(* IEC 61131-3 sources: daoli-st-library/DL_Device (part 14) *)

(* ---- FB_DL_BushingDrawStartSeq.st ---- *)
// FB_DL_BushingDrawStartSeq v1.0.0
// 开源溯源：clean-room 自研（族 DL_Device，ST 生态实测 0 命中，无外部代码引入）
(*
  功能: 拉丝启动八相顺控：IDLE→HEAT→(达标保持300s)DRIP→(检滴料)ATTACH→(丝根附着)RAMP
        →(达目标速度)STEADY→(断丝)BREAK→(重接)RAMP；RAMP 按 20 m/min² 斜坡（增量 (20/60)·fCycleS）。
        联锁：①HEAT 相温度未达 fTempTarget − 5 °C 前 xWinderEnable 必须 FALSE；
              ②BREAK 相速度降至 fSpeedTarget·0.3 并保持 60 s 等重接，超时锁存；
              ③FAULT 相 xWinderEnable = FALSE 且 fSpeedCmd = 0（安全侧），仅 xReset 解除。
  邻件: 与 FC_DL_BushingTempZoneCalc（分区温度）、FC_DL_BushingPowerBalanceCalc（功率平衡）同族，本件不调用 FC。
  码表: 9331 入参非有限｜9332 组态非法(fCycleS/fTempTarget/fSpeedTarget≤0)｜9333 相超时(1800/60/60/120/60 s)
        9334 相位落 ELSE 兜底｜9335 信息级进入稳态拉丝。故障码锁存至 xReset 上升沿。
  边界: 无方法块/无属性块/无全局变量/无物理 IO 地址；六 TON 单相独占且无条件刷新；速度单位统一 m/min。
*)
TYPE E_DL_DrawStartPhase :
(
    IDLE   := 0,        // 空闲：等启动指令 [-] / Idle, waiting start
    HEAT   := 10,       // 升温：漏板升到目标 − 5 °C 并保持 [-] / Heating bushing
    DRIP   := 20,       // 滴料：等玻璃液滴料 [-] / Waiting for drip
    ATTACH := 30,       // 附着：等丝根附着 [-] / Waiting for attachment
    RAMP   := 40,       // 升速：按 20 m/min² 升至目标 [-] / Ramping up
    STEADY := 50,       // 稳态：稳态拉丝 [-] / Steady drawing
    BREAK  := 60,       // 断丝：降速至 30% 待重接 [-] / Break, slow for re-attach
    FAULT  := 90        // 故障：锁存，仅复位沿可出 [-] / Fault latched
);
END_TYPE
FUNCTION_BLOCK FB_DL_BushingDrawStartSeq
VAR_INPUT
    xEnable         : BOOL := FALSE;    // 使能，FALSE 时冻结在 IDLE [-] / Enable gate
    xStart          : BOOL := FALSE;    // 启动指令，上升沿有效 [-] / Start rising edge
    xReset          : BOOL := FALSE;    // 复位，上升沿清故障锁存 [-] / Reset rising edge
    fBushingTemp    : REAL := 25.0;     // 漏板实测温度 [°C] / Measured bushing temperature [degC]
    fTempTarget     : REAL := 1250.0;   // 漏板目标温度 [°C]，域 > 0 / Target temperature [degC]
    xDripDetected   : BOOL := FALSE;    // 滴料检出反馈 [-] / Drip detected
    xStrandAttached : BOOL := FALSE;    // 丝根附着反馈 [-] / Strand attached
    fWinderSpeed    : REAL := 0.0;      // 卷绕实测线速 [m/min] / Measured winder speed [m/min]
    fSpeedTarget    : REAL := 900.0;    // 目标拉丝线速 [m/min]，域 > 0 / Target speed [m/min]
    xBreakDetected  : BOOL := FALSE;    // 断丝检出反馈 [-] / Break detected
    fCycleS         : REAL := 0.01;     // 任务周期 [s]，域 > 0 / Task cycle time [s]
END_VAR
VAR_OUTPUT
    ePhase        : E_DL_DrawStartPhase;    // 相位出口，段尾单点映射 [-] / Phase outlet
    xHeatEnable   : BOOL;                   // 漏板加热使能（仅 HEAT 相）[-] / Heat enable
    xWinderEnable : BOOL;                   // 卷绕使能（温度达标后）[-] / Winder enable
    fSpeedCmd     : REAL;                   // 线速指令 [m/min] / Speed command [m/min]
    xSteady       : BOOL;                   // 稳态标志（STEADY 相电平）[-] / Steady flag
    xFault        : BOOL;                   // 故障锁存标志 [-] / Fault latch flag
    uErrorId      : UDINT;                  // 事件码，0 = 无事件 / Event code
END_VAR
VAR
    tonHeat   : TON;                        // 温度达标保持窗 300 s，无条件刷新 / Temperature dwell
    tonHeatTo : TON;                        // 升温相总超时 1800 s，无条件刷新 / Heat timeout
    tonDrip   : TON;                        // 滴料相超时 60 s，无条件刷新 / Drip timeout
    tonAttach : TON;                        // 附着相超时 60 s，无条件刷新 / Attach timeout
    tonRamp   : TON;                        // 升速相超时 120 s，无条件刷新 / Ramp timeout
    tonBreak  : TON;                        // 断丝保持窗 60 s，无条件刷新 / Break hold window
    rtStart   : R_TRIG;                     // 启动沿实例，无条件刷新 / Start edge instance
    rtReset   : R_TRIG;                     // 复位沿实例，无条件刷新 / Reset edge instance
    _ePhase   : E_DL_DrawStartPhase := E_DL_DrawStartPhase.IDLE;    // 内部相位，CASE 唯一写入 / Internal phase
    _fSpeed   : REAL := 0.0;                // 速度斜坡内部量 [m/min] / Ramp speed [m/min]
    _bReady   : BOOL := FALSE;              // 温度达标判据 [-] / Temperature ready judgement
    _bFault   : BOOL := FALSE;              // 故障锁存位（锁存量，仅复位沿清）/ Latched fault bit
    _uFault   : UDINT := 16#0000;           // 故障码锁存（锁存量，仅复位沿清）/ Latched fault code
    _uInfo    : UDINT := 16#0000;           // 信息码，每拍重算 / Transient info code
END_VAR
// 段 0：定时器与沿实例无条件周期刷新（禁置于 IF/CASE 内，R7/R188）/ Unconditional refresh
rtStart(CLK := xStart);                                                     // 启动沿每拍必调 / Start edge
rtReset(CLK := xReset);                                                     // 复位沿每拍必调 / Reset edge
tonHeat(IN := (_ePhase = E_DL_DrawStartPhase.HEAT) AND (fBushingTemp >= (fTempTarget - 5.0)), PT := T#300S);
tonHeatTo(IN := (_ePhase = E_DL_DrawStartPhase.HEAT), PT := T#1800S);       // 升温总超时 / Heat timeout
tonDrip(IN := (_ePhase = E_DL_DrawStartPhase.DRIP), PT := T#60S);           // 滴料超时 / Drip timeout
tonAttach(IN := (_ePhase = E_DL_DrawStartPhase.ATTACH), PT := T#60S);       // 附着超时 / Attach timeout
tonRamp(IN := (_ePhase = E_DL_DrawStartPhase.RAMP), PT := T#120S);          // 升速超时 / Ramp timeout
tonBreak(IN := (_ePhase = E_DL_DrawStartPhase.BREAK), PT := T#60S);         // 断丝保持窗 / Break window
// 段 1：单拍量预清零（锁存量 _bFault/_uFault/_fSpeed 不入清单，R187）/ One-shot clear
_uInfo := 16#0000;                  // 信息码每拍重算 / Info code recomputed
_bReady := FALSE;                   // 温度达标判据缺省假 / Ready default false
// 段 2：非有限闸与组态域闸（归因唯一，逐因独立码，R190）/ Gate stage
IF (fBushingTemp <> fBushingTemp) OR (fTempTarget <> fTempTarget)
   OR (fWinderSpeed <> fWinderSpeed) OR (fSpeedTarget <> fSpeedTarget) OR (fCycleS <> fCycleS)
   OR (ABS(fBushingTemp) >= 3.0E38) OR (ABS(fTempTarget) >= 3.0E38)
   OR (ABS(fWinderSpeed) >= 3.0E38) OR (ABS(fSpeedTarget) >= 3.0E38) OR (ABS(fCycleS) >= 3.0E38) THEN
    _uFault := 16#0002_9331;        // 故障级：入参非有限 / Fault: non-finite input
    _bFault := TRUE;                // 置故障锁存（R45 配对）/ Set fault latch
END_IF
IF (fCycleS <= 1.0E-6) OR (fTempTarget <= 1.0E-6) OR (fSpeedTarget <= 1.0E-6) THEN
    _uFault := 16#0002_9332;        // 故障级：组态非法 / Fault: illegal configuration
    _bFault := TRUE;                // 置故障锁存（R45 配对）/ Set fault latch
END_IF
// 段 3：温度达标判据（HEAT 与 DRIP 共用，禁 EQUAL 比较）/ Temperature ready judgement
IF fBushingTemp >= (fTempTarget - 5.0) THEN
    _bReady := TRUE;                // 达目标 − 5 °C / Reached target minus margin
END_IF
// 段 4：复位沿（FAULT 唯一解除路径）/ Reset edge, only exit from fault
IF rtReset.Q THEN                   // rtReset.Q = 当拍量 / Reset edge per scan
    IF _ePhase = E_DL_DrawStartPhase.FAULT THEN
        _ePhase := E_DL_DrawStartPhase.IDLE;    // 故障相迁出回空闲 / Fault exits to idle
    END_IF
    _fSpeed := 0.0;                 // 斜坡量归零（锁存量解除）/ Ramp cleared on reset
    _bFault := FALSE;               // 清故障锁存位（仅此解除沿可清）/ Clear latched bit
    _uFault := 16#0000;             // 清故障锁存码（仅此解除沿可清）/ Clear latched code
END_IF
// 段 5：相位机（本拍合法事件优先于超时，R275）/ Phase machine
CASE _ePhase OF
E_DL_DrawStartPhase.IDLE:
    IF _bFault THEN
        _ePhase := E_DL_DrawStartPhase.FAULT;       // 聚合故障进故障相 / Enter fault
    ELSIF rtStart.Q AND xEnable THEN
        _fSpeed := 0.0;                             // 启动前进度清零 / Ramp reset on start
        _ePhase := E_DL_DrawStartPhase.HEAT;        // 进升温相 / Enter heat
    END_IF
E_DL_DrawStartPhase.HEAT:
    IF _bFault THEN
        _ePhase := E_DL_DrawStartPhase.FAULT;       // 故障优先 / Fault first
    ELSIF NOT xEnable THEN
        _ePhase := E_DL_DrawStartPhase.IDLE;        // 使能撤销回空闲 / Enable dropped
    ELSIF tonHeat.Q THEN
        _ePhase := E_DL_DrawStartPhase.DRIP;        // 达标保持 300 s：进滴料相 / Dwell done, drip
    ELSIF tonHeatTo.Q THEN
        _uFault := 16#0002_9333;                    // 故障级：升温相超时 / Heat timeout
        _bFault := TRUE;                            // 置故障锁存（R45 配对）/ Set latch
        _ePhase := E_DL_DrawStartPhase.FAULT;       // 进故障相 / Enter fault
    END_IF
E_DL_DrawStartPhase.DRIP:
    IF _bFault THEN
        _ePhase := E_DL_DrawStartPhase.FAULT;       // 故障优先 / Fault first
    ELSIF NOT xEnable THEN
        _ePhase := E_DL_DrawStartPhase.IDLE;        // 使能撤销回空闲（安全侧，R92 修）/ Enable dropped to IDLE
    ELSIF xDripDetected THEN
        _ePhase := E_DL_DrawStartPhase.ATTACH;      // 检出滴料：进附着相 / Drip seen, attach
    ELSIF tonDrip.Q THEN
        _uFault := 16#0002_9333;                    // 故障级：滴料相超时 / Drip timeout
        _bFault := TRUE;                            // 置故障锁存（R45 配对）/ Set latch
        _ePhase := E_DL_DrawStartPhase.FAULT;       // 进故障相 / Enter fault
    END_IF
E_DL_DrawStartPhase.ATTACH:
    IF _bFault THEN
        _ePhase := E_DL_DrawStartPhase.FAULT;       // 故障优先 / Fault first
    ELSIF NOT xEnable THEN
        _ePhase := E_DL_DrawStartPhase.IDLE;        // 使能撤销回空闲（安全侧，R92 修）/ Enable dropped to IDLE
    ELSIF xStrandAttached THEN
        _fSpeed := 0.0;                             // 升速前进度清零 / Reset ramp before spinning
        _ePhase := E_DL_DrawStartPhase.RAMP;        // 进升速相 / Enter ramp
    ELSIF tonAttach.Q THEN
        _uFault := 16#0002_9333;                    // 故障级：附着相超时 / Attach timeout
        _bFault := TRUE;                            // 置故障锁存（R45 配对）/ Set latch
        _ePhase := E_DL_DrawStartPhase.FAULT;       // 进故障相 / Enter fault
    END_IF
E_DL_DrawStartPhase.RAMP:
    IF _bFault THEN
        _ePhase := E_DL_DrawStartPhase.FAULT;       // 故障优先 / Fault first
    ELSIF NOT xEnable THEN
        _ePhase := E_DL_DrawStartPhase.IDLE;        // 使能撤销回空闲（安全侧，R92 修）/ Enable dropped to IDLE
    ELSIF xBreakDetected THEN
        _ePhase := E_DL_DrawStartPhase.BREAK;       // 升速中断丝：进断丝相 / Break during ramp
    ELSIF _fSpeed >= fSpeedTarget THEN
        _uInfo := 16#0002_9335;                     // 信息级：进入稳态拉丝 / Info: steady reached
        _ePhase := E_DL_DrawStartPhase.STEADY;      // 达目标：进稳态相 / Target reached
    ELSIF tonRamp.Q THEN
        _uFault := 16#0002_9333;                    // 故障级：升速相超时 / Ramp timeout
        _bFault := TRUE;                            // 置故障锁存（R45 配对）/ Set latch
        _ePhase := E_DL_DrawStartPhase.FAULT;       // 进故障相 / Enter fault
    END_IF
E_DL_DrawStartPhase.STEADY:
    IF _bFault THEN
        _ePhase := E_DL_DrawStartPhase.FAULT;       // 故障优先 / Fault first
    ELSIF NOT xEnable THEN
        _ePhase := E_DL_DrawStartPhase.IDLE;        // 使能撤销回空闲 / Enable dropped
    ELSIF xBreakDetected THEN
        _ePhase := E_DL_DrawStartPhase.BREAK;       // 断丝：进断丝相 / Break, go break
    END_IF
E_DL_DrawStartPhase.BREAK:
    IF _bFault THEN
        _ePhase := E_DL_DrawStartPhase.FAULT;       // 故障优先 / Fault first
    ELSIF NOT xEnable THEN
        _ePhase := E_DL_DrawStartPhase.IDLE;        // 使能撤销回空闲（安全侧，R92 修）/ Enable dropped to IDLE
    ELSIF xStrandAttached AND (NOT xBreakDetected) THEN
        _ePhase := E_DL_DrawStartPhase.RAMP;        // 重接成功回升速相 / Re-attached, ramp
    ELSIF tonBreak.Q THEN
        _uFault := 16#0002_9333;                    // 故障级：重接等待超时 / Re-attach timeout
        _bFault := TRUE;                            // 置故障锁存（R45 配对）/ Set latch
        _ePhase := E_DL_DrawStartPhase.FAULT;       // 进故障相 / Enter fault
    END_IF
E_DL_DrawStartPhase.FAULT:
    IF rtReset.Q THEN
        _ePhase := E_DL_DrawStartPhase.IDLE;        // 复位沿解除（段 4 已清锁存）/ Reset releases
    END_IF
ELSE
    _uFault := 16#0002_9334;                        // 故障级：非法相位兜底 / Illegal phase id
    _bFault := TRUE;                                // 置故障锁存（R45 配对）/ Set latch
    _ePhase := E_DL_DrawStartPhase.FAULT;           // 强制进故障相 / Force into fault
END_CASE
// 段 6：速度斜坡（增量 = (20/60)·fCycleS，禁阶跃；BREAK 独立降速）/ Speed ramp
IF (_ePhase = E_DL_DrawStartPhase.RAMP) THEN
    _fSpeed := _fSpeed + 20.0 / 60.0 * fCycleS;     // 斜坡升速 [m/min] / Ramp up
    IF _fSpeed > fSpeedTarget THEN
        _fSpeed := fSpeedTarget;                    // 不得越过目标 / No overshoot
    END_IF
ELSIF (_ePhase = E_DL_DrawStartPhase.STEADY) THEN
    _fSpeed := fSpeedTarget;                        // 稳态保持目标速度 / Hold target speed
ELSIF (_ePhase = E_DL_DrawStartPhase.BREAK) THEN
    _fSpeed := fSpeedTarget * 0.3;                  // 断丝相立即降至 30% / Drop to 30 percent
ELSE
    _fSpeed := 0.0;                                 // 其余相（含故障/空闲）速度零 / Other phases zero
END_IF
// 段 7：出口单点映射（名实双出口，R191；安全侧再硬清零）/ Outlet mapping
ePhase := _ePhase;                                  // 相位出口单点映射 / Phase outlet
IF (_ePhase = E_DL_DrawStartPhase.FAULT) OR _bFault THEN
    xHeatEnable := FALSE;                           // 故障侧加热硬零 / Fault heat hard zero
    xWinderEnable := FALSE;                         // 故障侧卷绕硬零 / Fault winder hard zero
    fSpeedCmd := 0.0;                               // 故障侧速度硬零 / Fault speed hard zero
    xSteady := FALSE;                               // 故障侧撤稳态 / Clear steady
    xFault := TRUE;                                 // 故障锁存回放 / Replay latched flag
    uErrorId := _uFault;                            // 故障码锁存回放 / Replay latched code
ELSE
    IF _ePhase = E_DL_DrawStartPhase.HEAT THEN
        xHeatEnable := TRUE;                        // 升温相加热使能 / Heat enable in phase
    ELSE
        xHeatEnable := FALSE;                       // 其余相不加热 / No heating
    END_IF
    IF _bReady AND (_ePhase <> E_DL_DrawStartPhase.IDLE) THEN
        xWinderEnable := TRUE;                      // 温度达标且非空闲才放行卷绕 / Winder allowed
    ELSE
        xWinderEnable := FALSE;                     // 温度未达标强制 FALSE / Winder forced off
    END_IF
    fSpeedCmd := _fSpeed;                           // 速度指令出口 / Speed command outlet
    IF _ePhase = E_DL_DrawStartPhase.STEADY THEN
        xSteady := TRUE;                            // 稳态相电平 / Steady phase level
    ELSE
        xSteady := FALSE;                           // 非稳态相清标志 / Not steady
    END_IF
    xFault := FALSE;                                // 无故障 / No fault
    uErrorId := _uInfo;                             // 信息码每拍重算 / Transient info code
END_IF
IF (fSpeedCmd <> fSpeedCmd) OR (ABS(fSpeedCmd) >= 3.0E38) OR (fSpeedCmd < 0.0) THEN
    fSpeedCmd := 0.0;                               // 出口复核失败回零速 / Outlet recheck zero
    xWinderEnable := FALSE;                         // 出口复核失败切卷绕 / Cut winder
    xFault := TRUE;                                 // 出口复核失败置故障 / Raise fault
    uErrorId := 16#0002_9331;                       // 故障级：出口非有限 / Fault: non-finite outlet
END_IF
END_FUNCTION_BLOCK

(* ---- FB_DL_BypassValveTrim.st ---- *)
(*
  FB_DL_BypassValveTrim  —  旁通阀供回水压差 PI 微调 / Bypass valve differential-pressure PI trim
  分类 Category : DL_Device
  码位 Code     : 16#03_2_09
  版本 Version  : 1.0.0
  溯源 Source   : ModPID 语义借鉴 · clean-room 实现，仅借分类/参数域/命名，未复制源码
  功能 Function : 1) 供/回水压差闭环 PI 微调（复用 FB_DL_PidController，阀位死区与限幅）；
                  2) 压差无效冻结输出保持末次阀位（跟踪回投）；
                  3) 阀位输出钳行程域并置饱和码。
  边界 Boundary : ① 两压力（压差合成源）任一无效冻结输出保持末次阀位；
                  ② 阀位输出钳行程域并置饱和标志；
                  ③ 死区带宽非法（<= 0 或倒置）出厂报码；
                  ④ PID 参数 Ti/Td = 0 按「关闭」语义不判非法（T2-5 参数域惯例）；
                  ⑤ 压差传感器量程 0 邻域防除零（换算分母域闸）；
                  ⑥ 输出三行同向：阀位微调 → 饱和标志 → 冻结标志。
  依赖 Depends  : FB_DL_PidController × 1（PI 调节，每拍无条件调用）

  码表 Error codes（本件子码步进 16#10，避让邻件码位）:
    16#0002_0309 故障级：组态非法（死区 <= 0 / 行程域倒置 / 量程 <= 0）
    16#0002_0319 故障级：相 ID 越界（枚举兜底路径）
    16#0002_0329 信息级：压差无效输出冻结 / 阀位饱和钳位（不置 bError）
*)

TYPE E_DL_BvtPhase :
(
    eIdle   := 0,  // 空闲（阀位回下限）/ Idle, valve at low limit
    eTrim   := 10, // PI 微调运行 / PI trim running
    eFrozen := 20, // 压差无效冻结 / Frozen by invalid DP
    eFault  := 90  // 组态故障锁定 / Configuration fault locked
);
END_TYPE

FUNCTION_BLOCK FB_DL_BypassValveTrim
VAR_INPUT
    bEnable       : BOOL;                           // 总使能，FALSE 阀位回下限 / Master enable
    bReset        : BOOL;                           // 复位，上升沿清组态故障 / Reset, clears fault
    fDpKpa        : REAL;                           // 供/回水压差实测 [kPa] / Measured DP [kPa]
    fDpSpKpa      : REAL := 25.0;                   // 压差设定 [kPa]，域 > 0 / DP setpoint [kPa]
    fKp           : REAL := 1.5;                    // 比例增益 [1] / Proportional gain [1]
    tTi           : TIME := T#20S;                  // 积分时间 [s]，T#0S = 关闭积分 / Integral time, T#0S = off
    tTd           : TIME := T#0S;                   // 微分时间 [s]，T#0S = 关闭微分 / Derivative time, T#0S = off
    fDeadbandKpa  : REAL := 0.5;                    // 控制死区 [kPa]，域 > 0 / Control deadband [kPa]
    fValveMinPct  : REAL := 0.0;                    // 阀位行程域下限 [%] / Valve domain low [%]
    fValveMaxPct  : REAL := 100.0;                  // 阀位行程域上限 [%] / Valve domain high [%]
    fManValvePct  : REAL := 50.0;                   // 手动阀位 [%]（跟踪回投基准）/ Manual valve position [%]
    fEps          : REAL := 1.0E-6;                 // 浮点判零容差 [1] / Floating zero tolerance
END_VAR
VAR_OUTPUT
    fValveOutPct  : REAL;                           // 旁通阀位输出 [%] / Bypass valve output [%]
    bSaturated    : BOOL;                           // 阀位饱和标志 / Valve saturated flag
    bFrozen       : BOOL;                           // 压差无效冻结标志 / Frozen by invalid DP
    bError        : BOOL;                           // 故障标志，与故障级码配对 / Fault flag
    uErrorId      : UDINT;                          // 事件码，0 = 无事件 / Event code
    eStateOut     : E_DL_BvtPhase;                  // 状态机当前态，段尾单点映射 / Phase mapped at tail
END_VAR
VAR
    _eState       : E_DL_BvtPhase := E_DL_BvtPhase.eIdle;  // 内部状态 / Internal state
    fbPid         : FB_DL_PidController;            // PI 实例（无条件调用）/ PI instance
    rtrReset      : R_TRIG;                         // 复位沿 / Reset edge
    bCfgOk        : BOOL;                           // 组态合法标志 / Configuration valid
    bDpOk         : BOOL;                           // 压差本拍有效 / DP valid this scan
    fValveHold    : REAL;                           // 末次有效阀位 [%]（冻结保持）/ Last valid valve position [%]
    uFault        : UDINT;                          // 锁存故障码 / Latched fault code
    uInfo         : UDINT;                          // 信息级码 / Information code
END_VAR

(* === 段 0 · 实例刷新 === *)
rtrReset(CLK := bReset);                          // 每拍刷新复位沿

(* === 段 1 · 组态闸（Ti/Td = 0 按「关闭」语义不判非法）=== *)
bCfgOk := (fDeadbandKpa > fEps)                   // 死区正域（<= 0 出厂报码）
          AND (fValveMaxPct > fValveMinPct + fEps)// 行程域不倒置
          AND (fDpSpKpa > fEps)                   // 设定正域
          AND (fDpSpKpa = fDpSpKpa) AND (fKp = fKp);  // NaN 自反（Ti/Td 为 0 合法：关闭语义）
IF NOT bCfgOk THEN
    uFault := 16#0002_0309;                       // 故障级：组态非法
END_IF
IF rtrReset.Q AND bCfgOk THEN
    uFault := 16#0000;                            // 复位沿清锁存（解除路径可达）
END_IF
uInfo := 16#0000;                                 // 信息码每拍清零
bDpOk := (fDpKpa = fDpKpa) AND (fDpKpa >= 0.0) AND (fDpKpa < 1.0E30);   // 压差 NaN 自反 + 非负域闸

(* === 段 2 · PI 实例（每拍无条件调用）=== *)
fbPid(bEnable := bEnable AND bCfgOk AND bDpOk,    // 压差无效/故障：PI 停调
      bManual := FALSE,                           // 自动微调
      fSetpoint := fDpSpKpa,                      // 压差设定
      fActual := fDpKpa,                          // 压差实测
      fKp := fKp,                                 // 比例增益
      tTi := tTi,                                 // 积分时间（0 = 关闭，合法语义）
      tTd := tTd,                                 // 微分时间（0 = 关闭）
      fDeadband := fDeadbandKpa,                  // 控制死区
      rOutMin := fValveMinPct,                    // 输出下限 = 行程域下限
      rOutMax := fValveMaxPct,                    // 输出上限 = 行程域上限
      tSampleTime := T#100MS,                     // 采样周期
      bTrack := (NOT bDpOk) OR (NOT bEnable),     // 无效/失能：跟踪回投保持阀位（无扰冻结）
      fTrackValue := fValveHold,                  // 跟踪值 = 末次有效阀位
      bReset := rtrReset.Q);                      // 复位沿透传

(* === 段 3 · 输出域闸与饱和标志 === *)
fValveOutPct := fbPid.fOut;                       // 阀位输出
IF fValveOutPct > fValveMaxPct THEN
    fValveOutPct := fValveMaxPct;                 // 钳到行程域上限
END_IF
IF fValveOutPct < fValveMinPct THEN
    fValveOutPct := fValveMinPct;                 // 钳到行程域下限
END_IF
bSaturated := fbPid.bLimitHigh OR fbPid.bLimitLow;   // 饱和标志（映射实例触限）
IF bSaturated AND bDpOk THEN
    uInfo := 16#0002_0329;                        // 信息级：阀位饱和钳位
END_IF

(* === 段 4 · 主状态机（ENUM + CASE，含 ELSE 兜底）=== *)
CASE _eState OF
E_DL_BvtPhase.eIdle :
    IF uFault <> 16#0000 THEN
        _eState := E_DL_BvtPhase.eFault;          // 故障优先
    ELSIF bEnable AND bCfgOk AND (NOT bDpOk) THEN
        _eState := E_DL_BvtPhase.eFrozen;         // 压差无效进冻结
    ELSIF bEnable AND bCfgOk AND bDpOk THEN
        _eState := E_DL_BvtPhase.eTrim;           // 进微调相
    END_IF

E_DL_BvtPhase.eTrim :
    IF (uFault <> 16#0000) OR (NOT bEnable) THEN
        _eState := E_DL_BvtPhase.eFault;          // 故障/失能转出
    ELSIF NOT bDpOk THEN
        uInfo := 16#0002_0329;                    // 信息级：压差无效输出冻结
        _eState := E_DL_BvtPhase.eFrozen;         // 转冻结相（阀位保持末次值）
    ELSE
        fValveHold := fValveOutPct;               // 有效拍记账末次阀位（冻结保持源）
    END_IF

E_DL_BvtPhase.eFrozen :
    IF bDpOk AND bEnable AND (uFault = 16#0000) THEN
        _eState := E_DL_BvtPhase.eTrim;           // 压差恢复回微调（解除路径可达，跟踪无扰）
    END_IF

E_DL_BvtPhase.eFault :
    IF uFault = 16#0000 THEN
        _eState := E_DL_BvtPhase.eIdle;           // 解锁回空闲
    END_IF

ELSE
    _eState := E_DL_BvtPhase.eFault;              // 非法状态拦截
    uFault := 16#0002_0319;                       // 故障级：相 ID 越界
END_CASE
bFrozen := (_eState = E_DL_BvtPhase.eFrozen);     // 冻结标志段尾单点映射

(* === 段 5 · 输出映射 === *)
bError := (uFault <> 16#0000);                    // 故障标志仅由故障级码置位（R45 配对）
IF bError THEN
    uErrorId := uFault;                           // 故障级优先上报
ELSE
    uErrorId := uInfo;                            // 否则上报信息级码
END_IF
eStateOut := _eState;                             // 输出枚举段尾单点映射（N2 规则）
END_FUNCTION_BLOCK

(* ---- FB_DL_CabinetCoolingWatch.st ---- *)
(*==============================================================================
 * 组件名称 (Component)  : FB_DL_CabinetCoolingWatch
 * 所属子库 (Sublibrary) : DL_Device
 * 当前版本 (Version)    : 1.0.0
 * 兼容性   (Platform)   : CODESYS 3.5 / TwinCAT 3 / 汇川 InoProShop / Machine Expert
 *                         仅依赖 Standard.library（TON / R_TRIG / TIME_TO_LREAL），零厂商方言
 * 来源标签 (Source)     : self-std
 * 功能描述 (Function)   : 控制柜热管理监视，三判据 -> NE107 降级出口：
 *                         ① 柜内-环境温差超限（热交换失效判据），确认窗满 ->
 *                            eMaintenanceReq；
 *                         ② 柜内风扇双判据（运行反馈缺失 OR 转速低于下限），
 *                            确认窗满 -> eCheckFunction；
 *                         ③ 滤网阻塞趋势——同环境温度下温差缓升速率（滑动窗
 *                            前后半均值斜率）超限 -> eMaintenanceReq。
 *                         只告警不控风扇：执行归调用方，本件零输出侧风扇操作
 *                         （「算一个值 / 做一件事」边界）。
 * 同类邻件互引 (Watch)  : 后缀 *Watch 族边界——触发 / 心跳类设备级监视归
 *                         FB_DL_CameraHealthWatch，时钟漂移类归 FB_DL_ClockDriftMonitor，
 *                         本件只负责热管理温差与风扇反馈域，三者互不替代。
 * 边界与语义披露 (Boundary disclosure) :
 *   1) 两温度非有限 -> 故障级锁存（各自独立码位，R190 归因唯一），健康出口
 *      eFailure（信号不可信）；解除路径 = 复位沿 AND 对应信号恢复有限。
 *   2) 环境温度高于柜内（温差 <= 0）为自然工况：判据挂起不发布、不计码
 *      （挂起态由 bJudgeSuspended 直接观测，R90 反证成立不加码）。
 *   3) 趋势窗样本数不足 nTrendWin 时趋势判据挂起（R307：挂起同步挂起累计载体
 *      ——样本只在监视中采集，挂起期不采不计）。
 *   4) 风扇转速反馈非有限 -> 故障级锁存（判据挂起 + eFailure）。
 *   5) 趋势样本仅在 ΔT > 0 时采集：负温差（环境更热）样本会稀释缓升斜率，
 *      滤网阻塞判据只对正温差域有意义。
 * 故障码表 (Error codes) :
 *   16#0003_050E [故障级] 柜内温度非有限，锁存，eFailure
 *                 反证：eFailure 不承载成因（三路信号三因，R190 必须码位互异）。
 *   16#0003_050F [故障级] 环境温度非有限，锁存，eFailure
 *                 反证：环温失效与柜温失效对健康出口同为 eFailure，组合不可区分。
 *   16#0003_0510 [故障级] 风扇转速反馈非有限，锁存，eFailure
 *                 反证：风扇反馈失效与两温度失效对健康出口同为 eFailure，组合不可区分。
 *   16#0003_0511 [故障级] 组态非法（确认窗 / 阈值域 / 趋势窗长 / 采样周期），已回退
 *                 反证：回退后监视继续，码位是组态错误唯一可见出口。
 *   16#0003_040A [信息级] 温差超限确认窗满（eMaintenanceReq 依据一）
 *                 反证：eHealth 为分级状态不承载成因；三判据三因码位互异（R190）。
 *   16#0003_040B [信息级] 风扇反馈失配确认窗满（eCheckFunction 依据）
 *                 反证：风扇失配分级（eCheckFunction）与温差成因分级（eMaintenanceReq）不同档，码位独立承载。
 *   16#0003_040C [信息级] 滤网阻塞趋势确认（eMaintenanceReq 依据二）
 *                 反证：趋势确认与温差确认同为 eMaintenanceReq 档，但成因互异，码位必须独立。
 * 码位总账 (Code ledger) : 16#0003_050E / 050F / 0510 / 0511 用 ｜ 16#0003_040A / 040B / 040C 用
 * 依赖     (Depends)    : TYPE E_DL_Ne107Status（属主 I_DL_DeviceHealth.st，只引用）
 * 红线自检 (Redline)    : R1 ✓ 零全局变量与 VAR_EXTERNAL ｜ R2 ✓ 零 %I/%Q 物理地址
 *                         R3 ✓ 纯 IEC 61131-3 ｜ R4 ✓ 非有限双判 / 斜率分母 eps 闸 / 域闸全枚举
 *                         R5 ✓ 全变量中英双语同行注释 ｜ R6 ✓ 三态 ENUM + CASE + ELSE 兜底
 *                         R7 ✓ 一沿二计时主体最前部无条件刷新
 * 修订历史 (Revision)   :
 *   2026-11-22  v1.0.0  首版入库（R68 构建轮 · 批 2 · 目标 11）
 *============================================================================*)

(*-----------------------------------------------------------------------------
 * 枚举: E_DL_CoolWatchState（归属 DL_Device，与 FB_DL_CabinetCoolingWatch 同文件）
 *----------------------------------------------------------------------------*)
TYPE E_DL_CoolWatchState :
(
    eIdle  := 0,    // 未使能：判据与趋势冻结 / Disabled, criteria and trend frozen
    eRun   := 10,   // 监视中：三判据并行评估 / Watching, three criteria evaluated
    eFault := 99    // 信号 / 组态锁存：判据挂起 / Signal or config latched, criteria suspended
);
END_TYPE

(*==============================================================================
 * 功能块: FB_DL_CabinetCoolingWatch
 * 调用约定: 每个扫描周期无条件调用一次。
 *============================================================================*)
FUNCTION_BLOCK FB_DL_CabinetCoolingWatch
VAR_INPUT
    fTempCab     : REAL;                 // 柜内温度 [℃] / Cabinet temperature [degC]
    fTempAmb     : REAL;                 // 环境温度 [℃] / Ambient temperature [degC]
    bFanRunCmd   : BOOL;                 // 风扇运行命令（只读判据输入）/ Fan run command, judgement input only
    bFanRunFb    : BOOL;                 // 风扇运行反馈 / Fan run feedback
    fFanSpeedFb  : REAL;                 // 风扇转速反馈 [rpm] / Fan speed feedback [rpm]
    fFanSpeedMin : REAL := 500.0;        // 风扇转速下限 [rpm] / Fan speed floor [rpm]
    fDtLimitK    : REAL := 15.0;         // 温差超限阈 [K] / Delta-T over-limit threshold [K]
    tConfirmDt   : TIME := T#60S;        // 温差确认窗 [s] / Delta-T confirmation window [s]
    tFanConfirm  : TIME := T#10S;        // 风扇失配确认窗 [s] / Fan mismatch confirmation window [s]
    fTrendLimit  : REAL := 2.0;          // 滤网阻塞趋势阈 [K/h] / Filter clogging trend threshold [K per h]
    tSample      : TIME := T#1M;         // 趋势采样周期 [min] / Trend sampling period [min]
    nTrendWin    : INT  := 12;           // 趋势窗样本数 [个]，域 4..16 且为偶数 / Trend window samples, 4..16 even
    bEnable      : BOOL := TRUE;         // 使能 / Enable
    bReset       : BOOL;                 // 上升沿：清除信号 / 组态锁存 / Rising edge: clear signal and config latches
END_VAR
VAR_OUTPUT
    eHealth         : E_DL_Ne107Status;  // NE107 健康出口 / NE107 health verdict
    fDtNow          : REAL;              // 当前温差 [K] / Current delta-T [K]
    bJudgeSuspended : BOOL;              // 判据挂起（自然温差 / 样本不足）/ Judge suspended, natural or insufficient
    bFanMismatch    : BOOL;              // 风扇失配确认（保持型）/ Fan mismatch confirmed, level held
    bTrendConfirmed : BOOL;              // 滤网阻塞趋势确认（保持型）/ Trend confirmed, level held
    fTrendSlope     : REAL;              // 当前趋势斜率 [K/h] / Current trend slope [K per h]
    bError          : BOOL;              // 故障标志（信号 / 组态锁存归并）/ Fault flag merged
    uErrorId        : UDINT;             // 故障码，0 = 无故障 / Error code, 0 = none
    eState          : E_DL_CoolWatchState; // 当前状态（供 HMI 诊断）/ Current state
END_VAR
VAR
    fbTrigReset   : R_TRIG;              // 复位沿检测实例 / Reset edge detector
    tonDt         : TON;                 // 温差确认窗计时实例 / Delta-T confirmation timer
    tonFan        : TON;                 // 风扇失配确认窗计时实例 / Fan mismatch confirmation timer
    tonSample     : TON;                 // 趋势采样周期（自复位）实例 / Trend sampling timer, self resetting
    eStateInt     : E_DL_CoolWatchState; // 主状态机内部当前态 / Internal state machine state
    fDtInt        : REAL;                // 温差内部副本 [K] / Internal delta-T
    bCabBad       : BOOL;                // 柜温非有限 / Cabinet temp non-finite
    bAmbBad       : BOOL;                // 环温非有限 / Ambient temp non-finite
    bFanSigBad    : BOOL;                // 风扇转速非有限 / Fan speed non-finite
    bCabLatch     : BOOL;                // 柜温失效锁存 / Cabinet latch
    bAmbLatch     : BOOL;                // 环温失效锁存 / Ambient latch
    bFanLatch     : BOOL;                // 风扇反馈失效锁存 / Fan feedback latch
    bCfgLatch     : BOOL;                // 组态故障锁存 / Config fault latch
    bCfgBad       : BOOL;                // 本拍组态非法 / Config illegal this scan
    bDtExceeds    : BOOL;                // 温差超限判据（挂起时 FALSE）/ Delta-T exceeds, FALSE when suspended
    bFanMismatchInt : BOOL;              // 风扇失配确认内部副本 / Internal fan mismatch
    bTrendConfInt : BOOL;                // 趋势确认内部副本 / Internal trend confirmed
    bTrendActive  : BOOL;                // 本拍趋势斜率可发布 / Trend slope publishable
    afDtRing      : ARRAY[0..15] OF REAL; // 趋势温差样本环形窗 [K] / Delta-T trend ring [K]
    nTrendWinEff  : INT;                 // 钳位后趋势窗长 [个] / Clamped trend window length
    nTrendWrite   : INT;                 // 趋势窗写指针 [0..15] / Trend ring write pointer
    nTrendFill    : INT;                 // 趋势窗有效样本数 [个] / Trend ring fill count
    fMeanOld      : REAL;                // 前半窗均值 [K] / Older half mean [K]
    fMeanNew      : REAL;                // 后半窗均值 [K] / Recent half mean [K]
    fHalfHours    : REAL;                // 半窗时长折算小时 [h] / Half window in hours [h]
    nHalf         : INT;                 // 半窗样本数 [个] / Half window sample count
    nI            : INT;                 // 遍历索引 / Loop index
    fSlope        : REAL;                // 斜率中间量 [K/h] / Slope intermediate
    fSpeedMinEff  : REAL;                // 钳位后转速下限 [rpm] / Clamped speed floor
    fDtLimEff     : REAL;                // 钳位后温差阈 [K] / Clamped delta-T threshold
    fTrendLimEff  : REAL;                // 钳位后趋势阈 [K/h] / Clamped trend threshold
    bErrorInt     : BOOL;                // 本拍故障置位累加（出口归并）/ Fault set accumulator
    bFirstScan    : BOOL := TRUE;        // 上电首扫标志 / First-scan flag
END_VAR
VAR CONSTANT
    DL_CW_WIN_MIN   : INT  := 4;      // 趋势窗长下限 [个] / Trend window floor
    DL_CW_WIN_MAX   : INT  := 16;     // 趋势窗长上限 [个]，与数组维度一致 / Trend window ceiling
    DL_CW_EPS       : REAL := 1.0E-6; // 斜率分母判零容差 [h] / Slope denominator epsilon [h]
    DL_CW_FIN_LIM   : REAL := 1.0E30; // REAL 有限幅值判界 / REAL finiteness bound
    DL_CW_HOUR_MS   : REAL := 3600000.0; // 小时毫秒换算常数 [ms/h] / Hours to milliseconds factor
END_VAR

(*------------------------------------------------------------------------------
 * 段 1｜无条件刷新区（红线 R7）：一沿三计时全部位于主体最前部
 *      Unconditional refresh: one edge and three timers at the very top
 *      tonSample 为周期窗自复位（IN 串 bEnable AND NOT 自身 Q，R188）
 *-----------------------------------------------------------------------------*)
fbTrigReset(CLK := bReset);

tonDt(IN := bDtExceeds, PT := tConfirmDt);
tonFan(IN := bFanRunCmd AND (NOT bFanSigBad)
        AND ((NOT bFanRunFb) OR (fFanSpeedFb < fSpeedMinEff)),   // 反馈失效时判据整体挂起 / Suspended on bad feedback
       PT := tFanConfirm);
tonSample(IN := bEnable AND (NOT tonSample.Q), PT := tSample);

(*------------------------------------------------------------------------------
 * 段 2｜上电首扫：趋势窗显式清零
 *      First-scan init: trend ring cleared explicitly
 *-----------------------------------------------------------------------------*)
IF bFirstScan THEN
    eStateInt := E_DL_CoolWatchState.eIdle;
    FOR nI := 0 TO 15 DO
        afDtRing[nI] := 0.0;     // 趋势窗显式清零 / Trend ring cleared
    END_FOR
    nTrendWrite := 0;
    nTrendFill  := 0;
    bFirstScan  := FALSE;
END_IF

(*------------------------------------------------------------------------------
 * 段 3｜每拍预清（FB32-1）：单拍标志，禁入锁存 / 快照
 *      Per-scan preset: single-scan flags only
 *-----------------------------------------------------------------------------*)
bErrorInt := FALSE;

(*------------------------------------------------------------------------------
 * 段 4｜非有限闸（R272 全枚举：三个测量 REAL 入参）+ 组态域闸（限值 / 窗长 / 周期）
 *      Non-finite gates over the three measurement inputs, plus the config gate
 *      解除路径（R152 自证）：复位沿 AND 对应信号恢复有限 / 组态改对
 *-----------------------------------------------------------------------------*)
bCabBad    := (fTempCab <> fTempCab) OR ((fTempCab - fTempCab) <> (fTempCab - fTempCab))
              OR (ABS(fTempCab) >= DL_CW_FIN_LIM);
bAmbBad    := (fTempAmb <> fTempAmb) OR ((fTempAmb - fTempAmb) <> (fTempAmb - fTempAmb))
              OR (ABS(fTempAmb) >= DL_CW_FIN_LIM);
bFanSigBad := (fFanSpeedFb <> fFanSpeedFb) OR ((fFanSpeedFb - fFanSpeedFb) <> (fFanSpeedFb - fFanSpeedFb))
              OR (ABS(fFanSpeedFb) >= DL_CW_FIN_LIM);

IF bCabBad THEN
    bCabLatch := TRUE;
    uErrorId  := 16#0003_050E;   // 故障级：柜温非有限 / Fault: cabinet temp non-finite
    bErrorInt := TRUE;
END_IF
IF bAmbBad THEN
    bAmbLatch := TRUE;
    uErrorId  := 16#0003_050F;   // 故障级：环温非有限 / Fault: ambient temp non-finite
    bErrorInt := TRUE;
END_IF
IF bFanSigBad THEN
    bFanLatch := TRUE;
    uErrorId  := 16#0003_0510;   // 故障级：风扇反馈非有限 / Fault: fan feedback non-finite
    bErrorInt := TRUE;
END_IF

bCfgBad := (tConfirmDt <= T#0S) OR (tFanConfirm <= T#0S) OR (tSample <= T#0S)
           OR (fDtLimitK <= 0.0) OR (fDtLimitK <> fDtLimitK)
           OR (fFanSpeedMin < 0.0) OR (fFanSpeedMin <> fFanSpeedMin)
           OR (fTrendLimit <= 0.0) OR (fTrendLimit <> fTrendLimit)
           OR (nTrendWin < DL_CW_WIN_MIN) OR (nTrendWin > DL_CW_WIN_MAX);

IF bCfgBad THEN
    bCfgLatch := TRUE;
    uErrorId  := 16#0003_0511;   // 故障级：组态非法 / Fault: config illegal
    bErrorInt := TRUE;
END_IF

(* 两级回退取值（R117）：非法参数钳回默认常量，服务不中断 *)
(* Two-level fallback values *)
IF (fFanSpeedMin < 0.0) OR (fFanSpeedMin <> fFanSpeedMin) THEN
    fSpeedMinEff := 500.0;       // 回退默认转速下限 / Fallback default floor
ELSE
    fSpeedMinEff := fFanSpeedMin;
END_IF
IF (fDtLimitK <= 0.0) OR (fDtLimitK <> fDtLimitK) THEN
    fDtLimEff := 15.0;           // 回退默认温差阈 / Fallback default threshold
ELSE
    fDtLimEff := fDtLimitK;
END_IF
IF (fTrendLimit <= 0.0) OR (fTrendLimit <> fTrendLimit) THEN
    fTrendLimEff := 2.0;         // 回退默认趋势阈 / Fallback default threshold
ELSE
    fTrendLimEff := fTrendLimit;
END_IF
IF (nTrendWin < DL_CW_WIN_MIN) OR (nTrendWin > DL_CW_WIN_MAX) THEN
    nTrendWinEff := 12;          // 回退默认窗长 / Fallback default window
ELSE
    nTrendWinEff := nTrendWin;
END_IF

(*------------------------------------------------------------------------------
 * 段 5｜温差判据（挂起语义）：环温 >= 柜温为自然工况，判据挂起不发布
 *      Delta-T criterion with suspension: ambient hotter means natural, suspended
 *-----------------------------------------------------------------------------*)
fDtInt := fTempCab - fTempAmb;
fDtNow := fDtInt;

bDtExceeds := (NOT bCabBad) AND (NOT bAmbBad)
              AND (fDtInt > fDtLimEff);      // 挂起（温差 <= 0）通过不置判据承载 / Suspension by not asserting

(*------------------------------------------------------------------------------
 * 段 6｜趋势采样与斜率（周期窗自复位 TON 到期拍采一个样本）
 *      Trend sampling and slope, one sample per self-resetting window tick
 *-----------------------------------------------------------------------------*)
bTrendActive := FALSE;
fSlope       := 0.0;

IF tonSample.Q AND (eStateInt = E_DL_CoolWatchState.eRun)
   AND (NOT bCabBad) AND (NOT bAmbBad) AND (fDtInt > 0.0) THEN
    afDtRing[nTrendWrite] := fDtInt;     // 正温差样本入环 / Positive delta-T sample into ring
    nTrendWrite := nTrendWrite + 1;
    IF nTrendWrite >= nTrendWinEff THEN
        nTrendWrite := 0;                // 显式回卷 / Explicit wrap
    END_IF
    IF nTrendFill < nTrendWinEff THEN
        nTrendFill := nTrendFill + 1;    // 填充推进 / Fill up
    END_IF
END_IF

IF nTrendFill >= nTrendWinEff THEN
    nHalf := nTrendWinEff / 2;           // 半窗样本数（窗长已组态为偶数域）/ Half count
    fMeanOld := 0.0;
    fMeanNew := 0.0;
    FOR nI := 0 TO (nHalf - 1) DO
        fMeanOld := fMeanOld + afDtRing[nI];              // 前半窗求和 / Older half sum
        fMeanNew := fMeanNew + afDtRing[nI + nHalf];      // 后半窗求和 / Recent half sum
    END_FOR
    fMeanOld := fMeanOld / UDINT_TO_REAL(DINT_TO_UDINT(nHalf));
    fMeanNew := fMeanNew / UDINT_TO_REAL(DINT_TO_UDINT(nHalf));
    fHalfHours := (TIME_TO_LREAL(tSample) * UDINT_TO_REAL(DINT_TO_UDINT(nHalf))) / DL_CW_HOUR_MS;
    IF fHalfHours > DL_CW_EPS THEN
        fSlope := (fMeanNew - fMeanOld) / fHalfHours;     // 缓升斜率 [K/h]，分母已闸 / Slope, guarded
        bTrendActive := TRUE;
        IF fSlope > fTrendLimEff THEN
            bTrendConfInt := TRUE;                        // 趋势确认（保持型）/ Trend confirmed
            uErrorId      := 16#0003_040C;                // 信息级：趋势确认 / Info: trend confirmed
        ELSIF fSlope <= fTrendLimEff THEN
            bTrendConfInt := FALSE;                       // 回落清除 / Clear on recovery
        END_IF
    END_IF
END_IF

(*------------------------------------------------------------------------------
 * 段 7｜主状态机（红线 R6）：ENUM + CASE + ELSE 兜底
 *      Main state machine with the mandatory ELSE fallback
 *-----------------------------------------------------------------------------*)
CASE eStateInt OF

    E_DL_CoolWatchState.eIdle:
        IF bEnable AND (NOT bCabLatch) AND (NOT bAmbLatch) AND (NOT bFanLatch) AND (NOT bCfgLatch) THEN
            eStateInt := E_DL_CoolWatchState.eRun;
        END_IF

    E_DL_CoolWatchState.eRun:
        IF bCabLatch OR bAmbLatch OR bFanLatch OR bCfgLatch OR (NOT bEnable) THEN
            eStateInt := E_DL_CoolWatchState.eFault;   // 任一锁存即挂起 / Any latch suspends
        END_IF

    E_DL_CoolWatchState.eFault:
        (* 解除路径（R152 自证可达）：复位沿 AND 全部锁存源已恢复 *)
        IF fbTrigReset.Q AND (NOT bCabBad) AND (NOT bAmbBad) AND (NOT bFanSigBad) AND (NOT bCfgBad) THEN
            bCabLatch := FALSE;
            bAmbLatch := FALSE;
            bFanLatch := FALSE;
            bCfgLatch := FALSE;
            uErrorId  := 16#0000_0000;
            eStateInt := E_DL_CoolWatchState.eIdle;
        END_IF

    ELSE
        eStateInt := E_DL_CoolWatchState.eFault;
        uErrorId  := 16#0003_0511;
        bErrorInt := TRUE;

END_CASE;

(*------------------------------------------------------------------------------
 * 段 8｜风扇失配确认消化（保持型）：确认窗满置位，命令撤销 / 反馈恢复回落清除
 *      Fan mismatch confirmation, level held, cleared on recovery
 *-----------------------------------------------------------------------------*)
IF tonFan.Q THEN
    bFanMismatchInt := TRUE;
    uErrorId        := 16#0003_040B;   // 信息级：风扇失配确认 / Info: fan mismatch confirmed
ELSIF (NOT bFanRunCmd) OR (bFanRunFb AND (NOT bFanSigBad) AND (fFanSpeedFb >= fSpeedMinEff)) THEN
    bFanMismatchInt := FALSE;          // 回落清除 / Clear on recovery
END_IF

(*------------------------------------------------------------------------------
 * 段 9｜输出单一出口（范式 P-05）：健康分级由三判据保持型派生
 *      Single output exit: health derived from the three level-held criteria
 *-----------------------------------------------------------------------------*)
bJudgeSuspended := (eStateInt <> E_DL_CoolWatchState.eRun)
                   OR (fDtInt <= 0.0)
                   OR (nTrendFill < nTrendWinEff);

IF eStateInt <> E_DL_CoolWatchState.eRun THEN
    eHealth := E_DL_Ne107Status.eUnknown;        // 未使能 / 锁存：未知（信号失效另见 eFailure 口径）
    IF bCabLatch OR bAmbLatch OR bFanLatch THEN
        eHealth := E_DL_Ne107Status.eFailure;    // 测量信号不可信 / Measurement untrusted
    END_IF
ELSIF bFanMismatchInt THEN
    eHealth := E_DL_Ne107Status.eCheckFunction;  // 风扇失配 / Fan mismatch
ELSIF bTrendConfInt OR tonDt.Q THEN
    eHealth := E_DL_Ne107Status.eMaintenanceReq; // 温差超限确认或趋势确认 / Delta-T confirmed or trend
    IF tonDt.Q THEN
        uErrorId := 16#0003_040A;                // 信息级：温差确认 / Info: delta-T confirmed
    END_IF
ELSE
    eHealth := E_DL_Ne107Status.eOk;             // 全判据通过 / All pass
END_IF

bFanMismatch    := bFanMismatchInt;
bTrendConfirmed := bTrendConfInt;
fTrendSlope     := fSlope;
bError          := bErrorInt OR (eStateInt = E_DL_CoolWatchState.eFault);
eState          := eStateInt;
END_FUNCTION_BLOCK

(* ---- FB_DL_CabinetTempDerate.st ---- *)
(*
    FB_DL_CabinetTempDerate —— 柜内温度降额（多点取最大 + 分级降额 + 失效保持超时报警）
    ------------------------------------------------------------------
    组件名称  : FB_DL_CabinetTempDerate
    分类      : DL_Device / ThermalManagement
    前缀      : FB_DL_
    版本      : 1.0.0
    溯源      : 借鉴点 —— 变频器 / 伺服驱动器热管理的通行策略：柜内多点测温取
                最大值作为判据（热点决定降额，平均值会掩盖局部过热）、按温度
                分级给出输出降额系数（0~1 的倍率，送上层限幅）、测温点失效时
                **保持末次有效值**并计时，超时仍无有效值才报警。
                诊断分级口径参考 NE 107 的「失效 / 超出规格 / 功能检查 / 维护」
                四级分类思想（本件对应「失效需保持 + 超时上报」）。
                clean-room 声明 —— 零代码行复制；分级判据、保持结构、码位与
                双语文档全部本件自有，仅使用 IEC 61131-3 标准库 TON / R_TRIG。
                许可证 —— 本件 MIT；来源标签 ne107 指公开诊断分类术语，
                标准文本不属代码，无许可继承。
    平台      : 纯 IEC 61131-3，CODESYS 3.5 / TwinCAT 3 / InoProShop / Machine Expert 通用
    作者      : 道莅代码库 · PLC编程专家（R70 构建轮 · 批 3 · N10）
    ------------------------------------------------------------------
    功能说明  : 一 逐点筛查：abSensOk 为 FALSE 或该点温度非有限 → 该点判为失效，
                   不参与取最大（失效点绝不当作 0 °C 参与，否则热点会被掩盖）。
                二 取最大：在有效点中取最大值 fMaxTemp；有效点数为 0 时
                   fMaxTemp 保持末次有效值（_fHoldMax），并启动失效计时。
                三 分级降额（判据自上而下，先到先得）：
                   fMaxTemp >= fT3 → eTier3 系数 fK3（降额最深）
                   fMaxTemp >= fT2 → eTier2 系数 fK2
                   fMaxTemp >= fT1 → eTier1 系数 fK1
                   否则 eNormal 系数 1.0
                   分级用 ENUM + CASE，含 ELSE 兜底（非法等级 → 回 eNormal 且置 0803）。
                   分级为「逐拍重算」，不带回差 —— 柜温降额关注安全侧，且上层
                   限幅链路本身有速率限制，故不在此处引入回差（口径写死）。
                四 失效报警：全点失效持续 tSensFault → 锁存 0802（故障级），
                   并把降额系数**压到最保守值 fK3**（失效时无法判明温度，
                   必须按最深降额处置，这是失效安全方向）。
                五 部分失效（有有效点但不足全部）：置信息级 0804，bError 保持 FALSE，
                   降额照常按有效点计算。
    错误码    : 16#0002_0801 组态非法（温度分级非单调 / 系数不在 (0,1] / 非有限），锁存 —— 故障级
                16#0002_0802 全部测温点失效超时（无法判明柜温），锁存 —— 故障级
                16#0002_0803 非法降额等级枚举（CASE ELSE 兜底），锁存 —— 故障级
                16#0002_0804 部分测温点失效（仍按有效点降额运行），不锁存 —— 信息级
    码位总账  : 0801 / 0802 / 0803 用（故障级，锁存回放）｜ 0804 用（信息级，每拍重算）
    状态机    : 降额等级 E_DL_CtdTier 四态，CASE 全覆盖 + ELSE 兜底。
                判据链为逐拍组合判据，无相驻留；失效计时由 TON 自持。
    边界与披露: 一 组态闸（R272 逐项点名）：fT1 < fT2 < fT3 严格单调；三个系数均在
                   (0.0, 1.0] 内且 fK3 <= fK2 <= fK1（降额随温度单调不增，反置会导致
                   高温反而给出更大系数，属致命组态错误）；六量全部纳入非有限闸；
                二 数组下标安全：全部 FOR 循环以常量 DL_CAB_N 为界（编译期确定），
                   本件无任何「以引脚值作下标」的访问；
                三 出口语义（R191 名实双出口）：fDerateK 与 eTier 同源（同一 CASE
                   分支内成对赋值，故系数与等级恒一致）；bSensorAlarm 与 0802 同源；
                四 失能（bEn = FALSE）：fDerateK 输出**最保守值 fK3**（失能不等于
                   允许满载，安全方向），fMaxTemp 保持末次有效值，eTier 回 eNormal，
                   锁存位不被失能清除（须 bReset 上升沿）；
                五 定时器 _tonSensFault 与沿实例 _rtReset 每周期无条件调用（规则 ⑦）；
                六 零全局变量、零 VAR_EXTERNAL、零物理地址、无除法。
    修订记录  : 2026-11-22 v1.0.0 首次入库（R70 构建轮 · 批 3 · N10）
*)
TYPE E_DL_CtdTier :
(
    eNormal := 0,   (* 正常，降额系数 = 1.0 / normal, the derating factor is one *)
    eTier1  := 10,  (* 一级降额（>= fT1）/ tier one, at or above fT1 *)
    eTier2  := 20,  (* 二级降额（>= fT2）/ tier two, at or above fT2 *)
    eTier3  := 30   (* 三级降额（>= fT3，最深）/ tier three, the deepest, at or above fT3 *)
);
END_TYPE

FUNCTION_BLOCK FB_DL_CabinetTempDerate
VAR_INPUT
    bEn        : BOOL := TRUE;             (* 使能，[标志] / the enable *)
    bReset     : BOOL := FALSE;            (* 故障复位（上升沿有效），[标志] / the fault reset, rising edge *)
    arTempC    : ARRAY[1..4] OF LREAL;     (* 四个柜内测温点温度，[°C] / four cabinet temperature readings *)
    abSensOk   : ARRAY[1..4] OF BOOL;      (* 四个测温点有效性（变送器级），[标志] / the per point validity *)
    fT1        : LREAL := 45.0;            (* 一级降额起判温度，[°C]，须 < fT2 / the tier one threshold *)
    fT2        : LREAL := 55.0;            (* 二级降额起判温度，[°C]，须 < fT3 / the tier two threshold *)
    fT3        : LREAL := 65.0;            (* 三级降额起判温度，[°C]，须 > fT2 / the tier three threshold *)
    fK1        : LREAL := 0.85;            (* 一级降额系数，[无量纲]，域 (0,1] / the tier one factor *)
    fK2        : LREAL := 0.70;            (* 二级降额系数，[无量纲]，域 (0,1] / the tier two factor *)
    fK3        : LREAL := 0.50;            (* 三级降额系数（亦为失效保守值），[无量纲]，域 (0,1] / the tier three factor *)
    tSensFault : TIME := T#30S;            (* 全点失效报警延时，[ms] / the all-points-failed alarm delay *)
END_VAR
VAR_OUTPUT
    fMaxTemp     : LREAL;                  (* 有效点中的最高柜温（失效时保持末次值），[°C] / the highest valid temperature *)
    fDerateK     : LREAL := 1.0;           (* 降额系数（输出倍率），[无量纲] / the derating factor *)
    eTier        : E_DL_CtdTier := E_DL_CtdTier.eNormal; (* 降额等级出口，[等级] / the derating tier outlet *)
    bSensorAlarm : BOOL;                   (* 全点失效超时报警（保持型），[标志] / the all sensors failed alarm *)
    bPartialFail : BOOL;                   (* 部分测温点失效，[标志] / some points have failed *)
    bBusy        : BOOL;                   (* 失效计时进行中，[标志] / the failure timer is running *)
    bValid       : BOOL;                   (* 出口可信（非锁存故障），[标志] / the outlets are trustworthy *)
    bError       : BOOL;                   (* 故障标志，故障级码时为 TRUE / the error flag, TRUE on fault level *)
    nErrCode     : UDINT;                  (* 错误码，0 = 正常 / the error id, 0 = ok *)
END_VAR
VAR
    _rtReset     : R_TRIG;                 (* 复位上升沿实例（无条件调用）/ the reset rising edge instance *)
    _tonSensFault : TON;                   (* 全点失效报警计时实例（无条件调用）/ the all sensors failed timer *)
    _bFault      : BOOL;                   (* 故障锁存位，仅 bReset 上升沿解除 / the latched fault bit *)
    _nCodeLatch  : UDINT;                  (* 锁存成因码，故障期回放 / the latched cause code *)
    _bCfgBad     : BOOL;                   (* 组态非法标志（逐拍重算）/ the configuration fault flag *)
    _bEnGood     : BOOL;                   (* 运行许可（使能且无锁存故障）/ the run permit *)
    _eTier       : E_DL_CtdTier := E_DL_CtdTier.eNormal; (* 降额等级寄存器，[等级] / the tier register *)
    _fMax        : LREAL;                  (* 本轮取最大中间量，[°C] / the maximum temporary *)
    _fHoldMax    : LREAL;                  (* 末次有效最高温度（失效保持量），[°C] / the last valid maximum *)
    _bHaveMax    : BOOL;                   (* 已获得过有效最高温度，[标志] / a valid maximum was seen *)
    _nValid      : INT;                    (* 有效测温点数，[个] / the number of valid points *)
    _i           : INT;                    (* 循环下标，[号] / the loop index *)
    _bPtBad      : BOOL;                   (* 单点失效判据结果，[标志] / the point failure verdict *)
    _fK          : LREAL;                  (* 本轮降额系数中间量，[无量纲] / the factor temporary *)
END_VAR
VAR CONSTANT
    DL_CAB_N     : INT := 4;               (* 测温点数（与数组声明同源），[个] / the point count matching the arrays *)
    DL_CAB_FMAX  : LREAL := 1.0E6;         (* 非有限筛查幅值上限，[°C] / the finiteness screening cap *)
    DL_CAB_KONE  : LREAL := 1.0;           (* 满载系数（正常等级），[无量纲] / the full load factor *)
END_VAR

// 段 1｜出口预置（R256 统一出口预置）/ segment 1, preset every outlet
fDerateK     := fK3;                       // 系数出口先置最保守值（安全缺省）/ preset the factor to the most conservative value
eTier        := E_DL_CtdTier.eNormal;      // 等级出口先置正常（段 8 覆盖）/ preset the tier to normal, overwritten in segment 8
bSensorAlarm := FALSE;                     // 全点失效报警预清零（真值在段 8 由锁存映射）/ preset the alarm false
bPartialFail := FALSE;                     // 部分失效标志预清零 / preset the partial flag false
bBusy        := FALSE;                     // 忙碌标志预清零 / preset the busy flag false
bValid       := FALSE;                     // 可用标志预置假，健康路径再置真 / preset valid false
bError       := FALSE;                     // 故障标志预清零 / preset the error flag false
nErrCode     := 0;                         // 错误码预置无错 / preset the code to zero
_nValid      := 0;                         // 有效点数预清零 / preset the valid count
_fMax        := 0.0;                       // 最大值中间量预置零 / preset the maximum temporary
_fK          := fK3;                       // 系数中间量预置最保守值 / preset the factor temporary

// 段 2｜沿实例与定时器无条件调用（规则 ⑦）/ segment 2, the reset edge and the timer
_rtReset(CLK := bReset);                   // 复位沿，每周期无条件刷新 / the reset edge, refreshed every scan

// 段 3｜复位解除：唯一可到达的清除边（R188）/ segment 3, the only latch release edge
IF _rtReset.Q THEN                         // 复位上升沿 / the reset rising edge
    _bFault     := FALSE;                  // 解除故障锁存 / release the fault latch
    _nCodeLatch := 0;                      // 清锁存码 / clear the latched code
END_IF

// 段 4｜组态守卫（R272 逐项点名，含单调性反置拦截）/ segment 4, the configuration guard
_bCfgBad := (fT1 >= fT2) OR (fT2 >= fT3)                                   // 温度分级非严格单调 / the tiers are not strictly monotonic
         OR (fK1 <= 0.0) OR (fK1 > DL_CAB_KONE)                            // 一级系数域外 / the tier one factor out of range
         OR (fK2 <= 0.0) OR (fK2 > DL_CAB_KONE)                            // 二级系数域外 / the tier two factor out of range
         OR (fK3 <= 0.0) OR (fK3 > DL_CAB_KONE)                            // 三级系数域外 / the tier three factor out of range
         OR (fK3 > fK2) OR (fK2 > fK1)                                     // 降额随温度反置（致命组态错）/ the factors increase with temperature
         OR (fT1 <> fT1) OR ((fT1 - fT1) <> 0.0) OR (ABS(fT1) > DL_CAB_FMAX)
         OR (fT2 <> fT2) OR ((fT2 - fT2) <> 0.0) OR (ABS(fT2) > DL_CAB_FMAX)
         OR (fT3 <> fT3) OR ((fT3 - fT3) <> 0.0) OR (ABS(fT3) > DL_CAB_FMAX)
         OR (fK1 <> fK1) OR ((fK1 - fK1) <> 0.0) OR (ABS(fK1) > DL_CAB_FMAX)
         OR (fK2 <> fK2) OR ((fK2 - fK2) <> 0.0) OR (ABS(fK2) > DL_CAB_FMAX)
         OR (fK3 <> fK3) OR ((fK3 - fK3) <> 0.0) OR (ABS(fK3) > DL_CAB_FMAX);

// 段 5｜首次成因锁存（故障期不重推断，R189）/ segment 5, the first cause latch
IF NOT _bFault THEN                        // 未锁存才登记 / register only while healthy
    IF _bCfgBad THEN                       // 组态非法 / an illegal configuration
        _bFault     := TRUE;               // 置锁存 / latch it
        _nCodeLatch := 16#0002_0801;       // 故障级：组态非法 / fault level: an illegal configuration
    END_IF
END_IF
_bEnGood := bEn AND NOT _bFault;           // 运行许可 / the run permit

// 段 6｜逐点筛查与取最大（常量上下界，下标安全）/ segment 6, the point screening and the maximum
_nValid := 0;                              // 有效点数清零重算 / recount the valid points
_fMax   := 0.0;                            // 最大值清零重算 / reset the maximum
FOR _i := 1 TO DL_CAB_N DO                 // 常量上下界 / constant bounds
    _bPtBad := (NOT abSensOk[_i])                                  // 变送器报失效 / the transmitter reports a failure
            OR (arTempC[_i] <> arTempC[_i])                        // NaN 自反判 / the NaN test
            OR ((arTempC[_i] - arTempC[_i]) <> 0.0)                // Inf 差值自反判 / the Inf test
            OR (ABS(arTempC[_i]) > DL_CAB_FMAX);                   // 幅值上界 / the amplitude cap
    IF NOT _bPtBad THEN                    // 有效点 / a valid point
        _nValid := _nValid + 1;            // 计数 / count it
        IF _nValid = 1 THEN                // 第一个有效点 / the first valid point
            _fMax := arTempC[_i];          // 直接作为当前最大 / take it as the maximum
        ELSIF arTempC[_i] > _fMax THEN     // 后续更大值 / a later larger value
            _fMax := arTempC[_i];          // 刷新最大 / refresh the maximum
        END_IF
    END_IF
END_FOR

// 段 7｜有效点处理：全失效保持 + 部分失效信息码 / segment 7, the validity handling
IF _nValid > 0 THEN                        // 存在有效点 / at least one valid point
    _fHoldMax := _fMax;                    // 刷新末次有效最高温度 / refresh the last valid maximum
    _bHaveMax := TRUE;                     // 标记已有有效值 / mark that a valid value exists
    IF _nValid < DL_CAB_N THEN             // 有有效点但不足全部 / some points failed
        bPartialFail := TRUE;              // 部分失效标志 / the partial failure flag
        nErrCode     := 16#0002_0804;      // 信息级：部分失效（不置 bError，R45）/ info level, no fault flag
    END_IF
ELSE                                       // 全部失效 / every point failed
    bPartialFail := FALSE;                 // 全失效时部分失效位不置（归因唯一，R190）/ clear the partial flag
END_IF

// 段 8｜失效计时器无条件调用与报警锁存 / segment 8, the failure timer and its latch
_tonSensFault(IN := (_nValid = 0), PT := tSensFault); // 全点失效计时，每周期无条件调用
bBusy := _bEnGood AND (_nValid = 0) AND NOT _tonSensFault.Q; // 失效计时进行中
IF _bEnGood AND (_nValid = 0) AND _tonSensFault.Q THEN       // 全点失效超时 / all points failed long enough
    IF NOT _bFault THEN                    // 首次判定才登记 / register the cause once
        _bFault     := TRUE;               // 置锁存 / latch it
        _nCodeLatch := 16#0002_0802;       // 故障级：全点失效 / fault level: every point failed
    END_IF
END_IF

// 段 9｜最高温度出口与降额分级（ENUM + CASE + ELSE 兜底）/ segment 9, the maximum outlet and the tiering
IF _bHaveMax THEN                          // 已有有效值 / a valid value exists
    fMaxTemp := _fHoldMax;                 // 输出末次有效最高温度（失效期保持）/ output the held maximum
ELSE                                       // 从未获得有效值 / no valid value yet
    fMaxTemp := 0.0;                       // 输出零值（初值语义，已在边界声明）/ output zero, the documented initial value
END_IF
IF _bEnGood THEN                           // 运行许可成立才参与分级 / grade only while the run permit holds
    IF fMaxTemp >= fT3 THEN                // 三级判据 / the tier three criterion
        _eTier := E_DL_CtdTier.eTier3;     // 三级 / tier three
    ELSIF fMaxTemp >= fT2 THEN             // 二级判据 / the tier two criterion
        _eTier := E_DL_CtdTier.eTier2;     // 二级 / tier two
    ELSIF fMaxTemp >= fT1 THEN             // 一级判据 / the tier one criterion
        _eTier := E_DL_CtdTier.eTier1;     // 一级 / tier one
    ELSE                                   // 低于一级判据 / under the tier one threshold
        _eTier := E_DL_CtdTier.eNormal;    // 正常 / normal
    END_IF
ELSE                                       // 失能或锁存故障 / disabled or latched
    _eTier := E_DL_CtdTier.eNormal;        // 等级回正常（系数由段 10 压到最保守值）/ the tier returns to normal, the factor is clamped below
END_IF
CASE _eTier OF
    E_DL_CtdTier.eNormal:                  // 正常等级 / the normal tier
        _fK := DL_CAB_KONE;                // 系数 1.0 / the factor is one
    E_DL_CtdTier.eTier1:                   // 一级降额 / tier one
        _fK := fK1;                        // 系数取一级值 / the tier one factor
    E_DL_CtdTier.eTier2:                   // 二级降额 / tier two
        _fK := fK2;                        // 系数取二级值 / the tier two factor
    E_DL_CtdTier.eTier3:                   // 三级降额 / tier three
        _fK := fK3;                        // 系数取三级值 / the tier three factor
    ELSE                                   // 非法枚举兜底（回安全等级 + 置码，规则 ⑥）/ the illegal enumeration guard
        _eTier      := E_DL_CtdTier.eNormal; // 回安全等级 / force the safe tier
        _fK         := fK3;                // 系数压到最保守值 / clamp the factor to the most conservative
        _bFault     := TRUE;               // 置锁存 / latch it
        _nCodeLatch := 16#0002_0803;       // 故障级：非法降额等级 / fault level: an illegal tier value
END_CASE

// 段 10｜出口映射（名实双出口同源，R191；故障 / 失效压最保守系数）/ segment 10, the outlet mapping
IF _bEnGood AND NOT _bFault THEN           // 健康运行 / healthy and running
    fDerateK := _fK;                       // 系数出口取分级结果 / the factor follows the tier
    bValid   := _bHaveMax OR (_nValid > 0); // 有有效值即出口可信 / trustworthy once a valid value exists
ELSE                                       // 失能或锁存故障 / disabled or latched
    fDerateK := fK3;                       // 压到最保守系数（失效安全方向）/ clamp to the most conservative factor
    bValid   := FALSE;                     // 出口不可信 / the outlets are not trustworthy
END_IF
eTier        := _eTier;                    // 等级出口 = 寄存器（与系数同源成对赋值）/ the tier outlet mirrors the register
bSensorAlarm := _bFault AND (_nCodeLatch = 16#0002_0802); // 报警位与 0802 同源 / the alarm shares the 0802 latch
bError       := _bFault;                   // 故障标志与锁存同源 / the fault flag shares the latch
nErrCode     := _nCodeLatch;               // 锁存码回放；无锁存时保留段 7 的信息级 0804 / replay the latch, keep the info code otherwise
IF _nCodeLatch = 0 THEN                    // 无锁存故障 / no latched fault
    IF _nValid > 0 AND _nValid < DL_CAB_N THEN // 部分失效仍在 / some points still failed
        nErrCode := 16#0002_0804;          // 信息级：部分失效 / info level, a partial failure
    END_IF
END_IF
END_FUNCTION_BLOCK

(* ---- FB_DL_CameraHealthWatch.st ---- *)
(*==============================================================================
 * 组件名称 (Component)  : FB_DL_CameraHealthWatch
 * 所属子库 (Sublibrary) : DL_Device
 * 当前版本 (Version)    : 1.0.1
 * 兼容性   (Platform)   : CODESYS 3.5 / TwinCAT 3 / 汇川 InoProShop / Machine Expert
 *                         仅依赖 Standard.library（TON / R_TRIG），零厂商方言
 * 来源标签 (Source)     : t1-5-tcopen（视觉设备健康看门狗语义，clean-room 编写）
 * 功能描述 (Function)   : 视觉相机设备健康看门狗，三判据独立确认窗：
 *                         ① 触发结果超时：触发发出后 tTrigTimeout 内无结果返回，
 *                            连续 nTimeoutTrips 次超时 -> eCheckFunction；
 *                         ② 心跳丢失：tHeartbeatWin 周期窗内无任何结果返回 ->
 *                            eCheckFunction（下一次结果返回即恢复）；
 *                         ③ NG 率滑动窗趋势：nNgWindow 环形窗内 NG 率超
 *                            fNgRateLimit 且 tNgConfirm 确认窗满 -> eMaintenanceReq。
 *                         样本数不足 nNgMinSamples 时 NG 判据挂起不发布
 *                         （挂起同步挂起确认计时器，R307）。
 * 统计语义次源 (Stats)  : NG 率滑动窗沿用 FB_DL_SignalStatistics 的环形窗统计语义
 *                         （次源参照，不实例化——该件为 REAL 值统计器，位样本
 *                         环形由本件自建，语义对齐不复制实现）。
 * 边界与语义披露 (Boundary disclosure) :
 *   1) 三判据各带独立确认窗（R13 三分类范式）：超时窗 = tTrigTimeout，心跳窗 =
 *      tHeartbeatWin，NG 确认窗 = tNgConfirm，互不复用。
 *   2) 同拍竞态（R275）：结果返回沿与超时 / 心跳到期同拍时，结果沿优先消化
 *      （IF / ELSIF 结构性优先），超时不计入 streak。
 *   3) NG 率分母（有效样本数）为 0 或低于下限时判据挂起：不发布、不计码、
 *      确认计时器不计时（挂起同步挂起累计载体 R307）。
 *   4) 使能撤销不置故障：只复位统计（streak / NG 窗 / 确认器），健康回 eUnknown。
 *   5) 组态非法两级回退（R117）：非法参数钳回默认常量，看门狗继续服务并置
 *      故障级码（组态错误必须可见，但监视不停摆）。
 * 配比约束 (Timing ratios) : tHeartbeatWin > tTrigTimeout（心跳窗必须宽于触发窗，
 *      否则每次触发超时都会连带心跳判据，双判据互相污染）。
 * 故障码表 (Error codes) :
 *   16#0003_0504 [故障级] 组态非法（窗长 / 样本数 / NG 率限域 / 配比），已两级回退
 *                 反证：回退后看门狗继续服务，eHealth 与合法组态时组合相同，
 *                 码位是组态错误唯一可见出口。
 *   16#0003_0402 [信息级] 触发超时连续 nTimeoutTrips 次达成（eCheckFunction 依据一）
 *                 反证：eHealth 为分级状态不承载成因；三类成因必须码位互异（R190）。
 *   16#0003_0403 [信息级] 心跳丢失确认（eCheckFunction 依据二）
 *                 反证：心跳丢失与触发超时对 eHealth 的影响同为 eCheckFunction，组合不可区分。
 *   16#0003_0404 [信息级] NG 率趋势确认（eMaintenanceReq 依据）
 *                 反证：NG 趋势的分级与 eCheckFunction 级两成因不同档，码位仍需独立承载。
 * 码位总账 (Code ledger) : 16#0003_0504 用 ｜ 16#0003_0402 / 0403 / 0404 用
 * 依赖     (Depends)    : TYPE E_DL_Ne107Status（属主 I_DL_DeviceHealth.st，只引用）
 * 红线自检 (Redline)    : R1 ✓ 零全局变量与 VAR_EXTERNAL ｜ R2 ✓ 零 %I/%Q 物理地址
 *                         R3 ✓ 纯 IEC 61131-3 ｜ R4 ✓ 域闸全枚举 / 两级回退 / 计数饱和
 *                         R5 ✓ 全变量中英双语同行注释 ｜ R6 ✓ 三态 ENUM + CASE + ELSE 兜底
 *                         R7 ✓ 三沿三计时主体最前部无条件刷新
 * 修订历史 (Revision)   :
 *   2026-11-22  v1.0.0  首版入库（R68 构建轮 · 批 2 · 目标 7）
 *   2026-11-22  v1.0.1  终审就地修①：组态锁存解除路径可达化（复位沿 + 组态改对即清锁存，原 eFault 相不可达）
 *============================================================================*)

(*-----------------------------------------------------------------------------
 * 枚举: E_DL_CamHealthState（归属 DL_Device，与 FB_DL_CameraHealthWatch 同文件）
 *----------------------------------------------------------------------------*)
TYPE E_DL_CamHealthState :
(
    eIdle  := 0,    // 未使能：统计复位，健康 eUnknown / Disabled, stats reset, eUnknown
    eWatch := 10,   // 监视中：三判据并行评估 / Watching, three criteria evaluated
    eFault := 99    // 组态故障：两级回退后继续监视 / Config fault, service continues after fallback
);
END_TYPE

(*==============================================================================
 * 功能块: FB_DL_CameraHealthWatch
 * 调用约定: 每个扫描周期无条件调用一次；结果引脚为单拍事件语义。
 *============================================================================*)
FUNCTION_BLOCK FB_DL_CameraHealthWatch
VAR_INPUT
    bTriggerOut     : BOOL;                 // 触发发出（上升沿登记未决）/ Trigger issued, rising edge arms outstanding
    bResultOk       : BOOL;                 // 本拍结果返回且 OK（单拍事件）/ Result returned OK this scan, single shot
    bResultNg       : BOOL;                 // 本拍结果返回且 NG（单拍事件）/ Result returned NG this scan, single shot
    tTrigTimeout    : TIME := T#5S;         // 触发结果超时窗 [s] / Trigger result timeout window [s]
    tHeartbeatWin   : TIME := T#30S;        // 心跳窗 [s]，须 > tTrigTimeout / Heartbeat window [s], must exceed trigger window
    tNgConfirm      : TIME := T#60S;        // NG 率确认窗 [s] / NG rate confirmation window [s]
    nTimeoutTrips   : INT  := 3;            // 连续超时次数阈值 [次] / Consecutive timeout trip threshold
    fNgRateLimit    : REAL := 0.2;          // NG 率上限 [1]，域 0..1 / NG rate ceiling, 0..1
    nNgMinSamples   : INT  := 5;            // NG 判据最小样本数 [个] / NG criterion minimum samples
    nNgWindow       : INT  := 32;           // NG 滑动窗长 [个]，域 2..64 / NG sliding window length
    bEnable         : BOOL := TRUE;         // 使能 / Enable
    bReset          : BOOL;                 // 上升沿：清组态故障锁存与统计 / Rising edge: clear config latch and stats
END_VAR
VAR_OUTPUT
    eHealth         : E_DL_Ne107Status;     // NE107 健康出口 / NE107 health verdict
    nTimeoutStreak  : INT;                  // 当前连续超时次数 [次] / Current consecutive timeout count
    bHeartbeatLost  : BOOL;                 // 心跳丢失（保持至下次结果）/ Heartbeat lost, held until next result
    fNgRate         : REAL;                 // 当前 NG 率 [1]，样本不足时为 -1.0 哨兵 / Current NG rate, -1.0 sentinel
    bNgSuspended    : BOOL;                 // NG 判据挂起（样本不足）/ NG criterion suspended, too few samples
    bError          : BOOL;                 // 故障标志（组态类锁存）/ Fault flag, configuration class
    uErrorId        : UDINT;                // 故障码，0 = 无故障 / Error code, 0 = none
    eState          : E_DL_CamHealthState;  // 当前状态（供 HMI 诊断）/ Current state for HMI diagnosis
END_VAR
VAR
    fbTrigTrig      : R_TRIG;               // 触发沿检测实例 / Trigger edge detector
    fbTrigResult    : R_TRIG;               // 结果返回沿检测实例 / Result edge detector
    fbTrigReset     : R_TRIG;               // 复位沿检测实例 / Reset edge detector
    tonTrig         : TON;                  // 触发超时计时实例 / Trigger timeout timer
    tonHb           : TON;                  // 心跳窗计时实例 / Heartbeat window timer
    tonNg           : TON;                  // NG 确认窗计时实例 / NG confirmation timer
    eStateInt       : E_DL_CamHealthState;  // 主状态机内部当前态 / Internal state machine state
    bTrigOutPrev    : BOOL;                 // TON 调用时刻的未决快照（同拍竞态判据）/ Outstanding snapshot at TON call time
    bResultAny      : BOOL;                 // 本拍有结果返回 / Any result this scan
    bTrigOutstanding: BOOL;                 // 触发未决（发出后未见结果）/ Trigger outstanding, no result yet
    bHbRun          : BOOL;                 // 心跳窗计时进行中 / Heartbeat window running
    bNgExceeds      : BOOL;                 // NG 率超限（挂起时强制 FALSE，驱动确认器）/ NG rate exceeds, drives the confirmer
    bNgConfirmed    : BOOL;                 // NG 判据已确认（保持型）/ NG criterion confirmed, level held
    abNgWin         : ARRAY[0..63] OF BOOL; // NG 样本环形窗（TRUE = NG）/ NG sample ring, TRUE = NG
    nNgWrite        : INT;                  // NG 窗写指针 [0..63] / NG ring write pointer
    nNgFill         : INT;                  // NG 窗有效样本数 [个] / NG ring valid samples
    nNgCount        : INT;                  // NG 窗内 NG 样本数 [个] / NG samples in ring
    nStreakInt      : INT;                  // 连续超时计数内部副本 / Internal timeout streak
    fNgRateInt      : REAL;                 // NG 率内部副本 [1] / Internal NG rate
    fNgLimEff       : REAL;                 // 钳位后 NG 率限 [1] / Clamped NG rate limit
    nWinEff         : INT;                  // 钳位后窗长 [个] / Clamped window length
    nMinEff         : INT;                  // 钳位后最小样本数 [个] / Clamped minimum samples
    nTripsEff       : INT;                  // 钳位后超时次数阈值 [次] / Clamped trip threshold
    bCfgBad         : BOOL;                 // 本拍组态非法 / Config illegal this scan
    bCfgLatch       : BOOL;                 // 组态故障锁存（复位沿清除）/ Config fault latch, cleared by reset edge
    bErrorInt       : BOOL;                 // 本拍故障置位累加（出口归并）/ Fault set accumulator of this scan
    bFirstScan      : BOOL := TRUE;         // 上电首扫标志 / First-scan flag
    nIdx            : INT;                  // 遍历索引 / Loop index
END_VAR
VAR CONSTANT
    DL_CH_WIN_MIN    : INT  := 2;     // NG 窗长下限 [个] / NG window floor
    DL_CH_WIN_MAX    : INT  := 64;    // NG 窗长上限 [个]，与数组维度一致 / NG window ceiling
    DL_CH_STREAK_MAX : INT  := 255;   // 超时计数饱和值 [次] / Timeout streak saturation
    DL_CH_RATE_NONE  : REAL := -1.0;  // NG 率不可发布哨兵 [1] / NG rate unpublishable sentinel
END_VAR

(*------------------------------------------------------------------------------
 * 段 1｜无条件刷新区（红线 R7）：三沿三计时全部位于主体最前部
 *      Unconditional refresh: three edges and three timers at the very top
 *      TON 的 IN 全部为内部派生量（R40 家族口径），禁挂外部引脚原值
 *-----------------------------------------------------------------------------*)
fbTrigTrig(CLK := bTriggerOut);
fbTrigResult(CLK := bResultOk OR bResultNg);
fbTrigReset(CLK := bReset);

tonTrig(IN := bTrigOutstanding, PT := tTrigTimeout);
tonHb(IN := bHbRun, PT := tHeartbeatWin);
tonNg(IN := bNgExceeds, PT := tNgConfirm);

(* 未决快照：取 TON 判定所依据的那一拍状态，供同拍竞态判据（R275） *)
(* Outstanding snapshot taken at TON call time for the same-scan race *)
bTrigOutPrev := bTrigOutstanding;

(*------------------------------------------------------------------------------
 * 段 2｜上电首扫：计数与环形窗显式清零，健康落 eUnknown
 *      First-scan init: counters and ring cleared, health to eUnknown
 *-----------------------------------------------------------------------------*)
IF bFirstScan THEN
    eStateInt := E_DL_CamHealthState.eIdle;
    eHealth   := E_DL_Ne107Status.eUnknown;
    FOR nIdx := 0 TO 63 DO
        abNgWin[nIdx] := FALSE;    // 环形窗显式清零 / Ring cleared explicitly
    END_FOR
    nNgWrite   := 0;
    nNgFill    := 0;
    nNgCount   := 0;
    nStreakInt := 0;
    fNgRateInt := DL_CH_RATE_NONE;
    bFirstScan := FALSE;
END_IF

(*------------------------------------------------------------------------------
 * 段 3｜每拍预清（FB32-1）：单拍标志，禁入锁存 / 快照
 *      Per-scan preset: single-scan flags only
 *-----------------------------------------------------------------------------*)
bErrorInt := FALSE;

(*------------------------------------------------------------------------------
 * 段 4｜组态域闸（R151 全枚举）+ 两级回退（R117）：非法钳回默认常量继续服务
 *      Config gate with two-level fallback: clamp to defaults, keep serving
 *      解除路径（R152 自证）：复位沿 AND 组态已改对
 *-----------------------------------------------------------------------------*)
bCfgBad := (tTrigTimeout <= T#0S) OR (tHeartbeatWin <= tTrigTimeout)
           OR (tNgConfirm <= T#0S) OR (nTimeoutTrips < 1)
           OR (nNgWindow < DL_CH_WIN_MIN) OR (nNgWindow > DL_CH_WIN_MAX)
           OR (nNgMinSamples < 1) OR (nNgMinSamples > nNgWindow)
           OR (fNgRateLimit < 0.0) OR (fNgRateLimit > 1.0) OR (fNgRateLimit <> fNgRateLimit);

IF bCfgBad THEN
    bCfgLatch := TRUE;
END_IF

(* 终审就地修 v1.0.1（R68）：解除路径（R152 自证可达）——复位沿 AND 组态非法条件
 * 全部消失即清锁存。原实现把锁存清零只写在 eFault 相分支，而组态闸置锁存后
 * 并不迁相至 eFault（只回 eIdle / 驻留），eFault 相不可达 -> 锁存永不可解，
 * 组件保护/监视功能一次性永久失效直至 PLC 重启（终审两式①）。
 * Clear path made provably reachable: reset edge with the illegal config gone. *)
IF fbTrigReset.Q AND (NOT bCfgBad) THEN
    bCfgLatch := FALSE;           // 锁存解除 / Latch cleared
    uErrorId  := 16#0000_0000;    // 码位随解除归零 / Code cleared with the latch
END_IF

(* 两级回退取值（非法值钳回默认常量，服务不中断） *)
(* Two-level fallback values, clamped to defaults, service continues *)
IF (fNgRateLimit < 0.0) OR (fNgRateLimit > 1.0) OR (fNgRateLimit <> fNgRateLimit) THEN
    fNgLimEff := 1.0;            // 回退默认：上限 1（判据退化为不触发）/ Fallback: no-trip ceiling
ELSE
    fNgLimEff := fNgRateLimit;   // 合法直通 / Valid pass-through
END_IF

IF (nNgWindow < DL_CH_WIN_MIN) OR (nNgWindow > DL_CH_WIN_MAX) THEN
    nWinEff := 32;               // 回退默认窗长 / Fallback default window
ELSE
    nWinEff := nNgWindow;        // 合法直通 / Valid pass-through
END_IF

IF (nNgMinSamples < 1) OR (nNgMinSamples > nWinEff) THEN
    nMinEff := 5;                // 回退默认最小样本 / Fallback default minimum
ELSE
    nMinEff := nNgMinSamples;    // 合法直通 / Valid pass-through
END_IF

IF nTimeoutTrips < 1 THEN
    nTripsEff := 1;              // 回退：单次超时即计 / Fallback: single trip counts
ELSE
    nTripsEff := nTimeoutTrips;  // 合法直通 / Valid pass-through
END_IF

IF bCfgLatch THEN
    uErrorId  := 16#0003_0504;   // 故障级：组态非法已回退 / Fault: config illegal, fallback applied
    bErrorInt := TRUE;           // R45 配对 / Paired with the fault code
END_IF

(*------------------------------------------------------------------------------
 * 段 5｜NG 率窗口统计（每拍重算）：写指针 / 样本数 / NG 计数 / 率
 *      NG ring statistics recomputed every scan
 *      挂起判据（R307）：有效样本数 < nMinEff 时 bNgExceeds 强制 FALSE（确认器停摆）
 *-----------------------------------------------------------------------------*)
bNgExceeds := FALSE;
fNgRateInt := DL_CH_RATE_NONE;

IF nNgFill >= nMinEff THEN
    fNgRateInt := UDINT_TO_REAL(DINT_TO_UDINT(nNgCount)) / UDINT_TO_REAL(DINT_TO_UDINT(nNgFill));  // 除子已闸 / Guarded denominator
    bNgSuspendedCalc := FALSE;   // 非挂起（占位变量见下方统一赋值）/ Not suspended, unified below
    IF fNgRateInt > fNgLimEff THEN
        bNgExceeds := TRUE;      // 超限（确认器计时窗口）/ Exceeds, confirmer timing
    END_IF
END_IF

(*------------------------------------------------------------------------------
 * 段 6｜主状态机（红线 R6）：ENUM + CASE + ELSE 兜底
 *      Main state machine with the mandatory ELSE fallback
 *      同拍竞态（R275）：结果沿优先于超时 / 心跳到期（IF / ELSIF 结构性优先）
 *-----------------------------------------------------------------------------*)
CASE eStateInt OF

    E_DL_CamHealthState.eIdle:
        IF bEnable AND (NOT bCfgLatch) THEN
            eStateInt := E_DL_CamHealthState.eWatch;
            bHbRun    := TRUE;           // 入监视相即立心跳窗（从未返回结果也可判丢失）/ Arm heartbeat on entry
        END_IF

    E_DL_CamHealthState.eWatch:
        IF bCfgLatch OR (NOT bEnable) THEN
            eStateInt := E_DL_CamHealthState.eIdle;
        ELSE
            (* —— ① 结果沿（最高优先）或超时到期，二者同拍时结果胜（R275） —— *)
            (* Result edge outranks the timeout expiry in the same scan *)
            IF fbTrigResult.Q THEN
                bTrigOutstanding := FALSE;
                nStreakInt  := 0;
                bHbRun      := TRUE;
                bHeartbeatLost := FALSE;
                abNgWin[nNgWrite] := bResultNg;    // NG 样本入环 / NG sample into ring
                nNgWrite := nNgWrite + 1;
                IF nNgWrite >= nWinEff THEN
                    nNgWrite := 0;                 // 显式回卷 / Explicit wrap
                END_IF
                IF nNgFill < nWinEff THEN
                    nNgFill := nNgFill + 1;        // 填充推进 / Fill up
                ELSE
                    IF abNgWin[nNgWrite] THEN      // 覆盖前扣减最旧样本的 NG 贡献 / Decrement the oldest
                        nNgCount := nNgCount - 1;
                    END_IF
                END_IF
                IF bResultNg THEN
                    nNgCount := nNgCount + 1;      // NG 计数推进 / NG count up
                END_IF
            ELSIF tonTrig.Q AND bTrigOutPrev THEN
                (* 超时消化：以 TON 判定拍的未决快照为准，不吞新触发沿 *)
                (* Timeout consumed against the snapshot, never eats a new trigger *)
                bTrigOutstanding := FALSE;
                IF nStreakInt < DL_CH_STREAK_MAX THEN
                    nStreakInt := nStreakInt + 1;  // 计数推进（饱和）/ Streak up, saturating
                END_IF
                IF nStreakInt >= nTripsEff THEN
                    uErrorId := 16#0003_0402;      // 信息级：超时三连 / Info: timeout streak
                END_IF
            END_IF

            (* —— ② 触发沿独立消化（与上段并行，不互斥） —— *)
            (* Trigger edge digested independently *)
            IF fbTrigTrig.Q THEN
                bTrigOutstanding := TRUE;
            END_IF

            (* —— ③ 心跳到期：置丢失（结果沿已优先重立心跳窗） —— *)
            (* Heartbeat expiry: lost flag set, result edge re-arms first *)
            IF bHbRun AND tonHb.Q THEN
                bHbRun         := FALSE;
                bHeartbeatLost := TRUE;
                uErrorId       := 16#0003_0403;   // 信息级：心跳丢失 / Info: heartbeat lost
            END_IF

            (* —— ④ NG 确认：超限确认窗满 -> 保持型确认（挂起时 bNgExceeds 已 FALSE） —— *)
            (* NG confirmation: confirmed level when the window fills *)
            IF tonNg.Q THEN
                bNgConfirmed := TRUE;
                uErrorId     := 16#0003_0404;     // 信息级：NG 趋势确认 / Info: NG trend confirmed
            ELSIF NOT bNgExceeds THEN
                bNgConfirmed := FALSE;            // 回落清除 / Clear on recovery
            END_IF
        END_IF

    E_DL_CamHealthState.eFault:
        (* 兜底态：解除路径 = 复位沿 AND 组态已改对（R152） *)
        IF fbTrigReset.Q AND (NOT bCfgBad) THEN
            bCfgLatch := FALSE;
            uErrorId  := 16#0000_0000;
            eStateInt := E_DL_CamHealthState.eIdle;
        END_IF

    ELSE
        (* 非法状态拦截：直接迁入兜底态并复用组态码（不隐式恢复） *)
        eStateInt := E_DL_CamHealthState.eFault;
        uErrorId  := 16#0003_0504;
        bErrorInt := TRUE;

END_CASE;

(*------------------------------------------------------------------------------
 * 段 7｜使能撤销复位统计（不置故障，规格明示）
 *      Enable withdrawal resets statistics without any fault
 *-----------------------------------------------------------------------------*)
IF (NOT bEnable) OR fbTrigReset.Q THEN
    nStreakInt := 0;             // 超时计数复位 / Streak reset
    nNgFill    := 0;             // 样本数复位 / Sample count reset
    nNgCount   := 0;             // NG 计数复位 / NG count reset
    nNgWrite   := 0;             // 写指针复位 / Write pointer reset
    bNgConfirmed := FALSE;       // NG 确认复位 / NG confirmation reset
    bHeartbeatLost := FALSE;     // 心跳丢失复位 / Heartbeat lost reset
    bTrigOutstanding := FALSE;   // 未决复位 / Outstanding reset
    bHbRun     := FALSE;         // 心跳窗复位 / Heartbeat window reset
END_IF

(*------------------------------------------------------------------------------
 * 段 8｜输出单一出口（范式 P-05）：健康分级由三判据保持型派生
 *      Single output exit: health derived from the three level-held criteria
 *-----------------------------------------------------------------------------*)
nTimeoutStreak := nStreakInt;
fNgRate := fNgRateInt;
bNgSuspended := (nNgFill < nMinEff);

IF (eStateInt = E_DL_CamHealthState.eIdle) OR (eStateInt = E_DL_CamHealthState.eFault) THEN
    eHealth := E_DL_Ne107Status.eUnknown;        // 未使能 / 故障：未知 / Idle or fault: unknown
ELSIF bNgConfirmed THEN
    eHealth := E_DL_Ne107Status.eMaintenanceReq; // NG 趋势确认 / NG trend confirmed
ELSIF (nStreakInt >= nTripsEff) OR bHeartbeatLost THEN
    eHealth := E_DL_Ne107Status.eCheckFunction;  // 超时三连或心跳丢失 / Streak or heartbeat lost
ELSE
    eHealth := E_DL_Ne107Status.eOk;             // 全判据通过 / All criteria pass
END_IF

bError := bErrorInt OR (eStateInt = E_DL_CamHealthState.eFault);
eState := eStateInt;
END_FUNCTION_BLOCK

(* ---- FB_DL_CartonErectVacMonitor.st ---- *)
(*
  FB_DL_CartonErectVacMonitor  —  纸箱成型吸盘真空建立时长与老化漂移监视 / Carton erector vacuum build-time and ageing monitor
  分类 Category : DL_Device
  码位 Code     : 16#03_2_10
  版本 Version  : 1.0.0
  来源 Source   : t2-1-lgf-measurement — IEC 61131-3 标准语义的道莅防御性实现
  溯源 Origin   : LGF 测量类文档公开语义借鉴（基线/漂移/样本中值），clean-room 实现，未复制源码行
  功能 Function : 1) 每次取料（bPickStart 上升沿）启动一次真空建立计时，真空度（负压绝对值）达 fVacTargetKpa
                     即记录本次建立时长 fBuildTimeMs；超 tBuildMax 未达则置 bBuildTimeout；
                  2) 建立时长入环形样本缓冲（长度 DL_BASE_MAX），基线 fBaselineMs 取**中值**（抗野值）；
                  3) 当前时长相对基线的漂移 fDriftPct 超 fDriftWarnPct 且连续 nWarnCycles 次 → bAgingWarn（吸盘老化）；
                  4) 样本数 < DL_MIN_SAMPLES 时不出漂移结论：bAgingWarn := FALSE、fDriftPct := 0（R191 显式声明）。
  边界 Boundary : ① fVacTargetKpa <= 0 判组态错 0210（建立判据门限为 0 会让"建立"恒成立）；
                      tBuildMax <= 0 / fDriftWarnPct <= 0 / nWarnCycles < 1 同判组态错；
                  ② nBaselineSamples > DL_BASE_MAX 时钳制到 DL_BASE_MAX 并置信息级 0110（不静默截断）；
                  ③ 建立时长为 0（同拍达成，或计时分辨率不足）走下限保护：分母用 MAX(基线, 1 ms)，
                     基线未建立（= 0）时 fDriftPct 直接置 0，绝不产生 inf/NaN；
                  ④ bBuildTimeout 为保持型（故障级 0220），清除路径 = rtReset.Q 或「下一次取料建立成功」；
                  ⑤ bAgingWarn 为维护级告警（信息级 0130，**不置 bError**）：漂移回落至门限内即自行释放；
                  ⑥ 注入件故障（iVac.bFault）时本件照常计时但置信息级 0140 并抑制漂移结论（数据不可信，
                     不得把注入件故障记成吸盘老化，R190 归因唯一）。
  依赖 Depends  : I_DL_VacuumGenerator（DL_Device 既有契约，注入不实例化）；
                  仅 Standard.library（TON / R_TRIG / ABS / MIN / MAX）
  同拍双窗配比  : tBuildMax（单次建立上限）与心跳窗 DL_HEART_WINDOW 不同源；配比约束
                  tBuildMax >= DL_HEART_WINDOW，保证建立过程中至少一次判活（R100）

  码表 Error codes（本件格 03_2_10，子码步进 +0x10）:
    16#0003_0210 故障级：组态非法（真空目标 <= 0 / 建立上限 <= 0 / 漂移门限 <= 0 / 预警次数 < 1）
    16#0003_0220 故障级：真空建立超时（tBuildMax 内未达 fVacTargetKpa，保持型）
    16#0003_0230 故障级：状态机落 ELSE 兜底（非法相位 ID）
    16#0003_0110 信息级：nBaselineSamples 超数组上限已钳制（不置 bError）
    16#0003_0120 信息级：样本数不足，本拍不出漂移结论（不置 bError）
    16#0003_0130 信息级：吸盘老化预警已成立（维护级，不置 bError）
    16#0003_0140 信息级：注入件故障，漂移结论抑制（不置 bError）

  修订历史 Revision :
    2026-11-18  v1.0.0  R37 首版
*)

TYPE E_DL_VacBuildState :
(
    eIdle    := 0,   // 空闲：等取料触发 / Idle, waiting for a pick trigger
    eBuilding := 10, // 建立中：本次真空建立计时进行中 / Building, timing the present evacuation
    eMeasured := 20, // 已测量：本次入样本缓冲，等下一次 / Measured, the sample is buffered
    eFault   := 90   // 故障：组态非法或建立超时锁定 / Fault, illegal configuration or a latched build timeout
);
END_TYPE

FUNCTION_BLOCK FB_DL_CartonErectVacMonitor
VAR_INPUT
    bEnable        : BOOL := FALSE;             // 总使能，FALSE 时不启动计时 / Master enable, low level stops timing
    bReset         : BOOL := FALSE;             // 复位，上升沿清故障锁存 / Reset, rising edge clears the latch
    bPickStart     : BOOL := FALSE;             // 取料起始触发（上升沿受理）/ Pick trigger, rising edge
    fVacTargetKpa  : REAL := 60.0;              // 真空目标（负压绝对值）[kPa]，域 > 0 / Vacuum target magnitude [kPa]
    tBuildMax      : TIME := T#1500MS;          // 单次建立时长上限 [ms]，域 > 0 / Maximum build time [ms]
    nBaselineSamples : INT := 9;                // 基线样本数 [个]，域 3~DL_BASE_MAX / Baseline sample count
    fDriftWarnPct  : REAL := 30.0;              // 漂移预警门限 [%]，域 > 0 / Drift warning threshold [%]
    nWarnCycles    : INT := 3;                  // 连续超门限次数 [次]，域 >= 1 / Consecutive exceed cycles
END_VAR
VAR_OUTPUT
    fBuildTimeMs   : REAL;                      // 本次建立时长 [ms] / Build time of the present pick [ms]
    fBaselineMs    : REAL;                      // 基线建立时长（样本中值）[ms] / Baseline build time, the sample median [ms]
    fDriftPct      : REAL;                      // 相对基线漂移 [%]，已限幅 / Drift against the baseline [%], clamped
    bAgingWarn     : BOOL;                      // 吸盘老化预警（维护级）/ Suction-cup ageing warning
    bBuildTimeout  : BOOL;                      // 建立超时（保持型）/ Build timeout, held
    nSampleCount   : INT;                       // 当前有效样本数 [个] / Number of valid samples
    bValid         : BOOL;                      // 判据可用标志 / Criteria usable
    bError         : BOOL;                      // 故障标志，派生自锁存 / Fault flag derived from the latch
    nErrId         : UDINT;                     // 事件码，0 = 无事件 / Event code, 0 = no event
    eStateOut      : E_DL_VacBuildState;        // 状态出口，段尾单点映射 / State outlet, mapped at the tail
END_VAR
VAR_IN_OUT
    iVac           : I_DL_VacuumGenerator;      // 真空发生器接口引用（注入，不实例化）/ Vacuum generator reference, injected
END_VAR
VAR
    tonBuild     : TON;                         // 单次建立计时，每拍无条件调用 / Build timer, called unconditionally
    tonHeart     : TON;                         // 周期心跳窗，自复位 / Periodic heartbeat window, self-resetting
    rtReset      : R_TRIG;                      // 复位上升沿 / Reset rising edge
    rtPick       : R_TRIG;                      // 取料上升沿 / Pick rising edge
    _eState      : E_DL_VacBuildState := E_DL_VacBuildState.eIdle;  // 内部相位（CASE 唯一写入目标）/ Internal phase
    _uFault      : UDINT;                       // 故障码锁存 / Latched fault code
    _uInfo       : UDINT;                       // 信息码，每拍重算 / Information code, recomputed per scan
    _bFault      : BOOL;                        // 故障锁存位 / Latched fault bit
    _bCfgBad     : BOOL;                        // 组态非法聚合 / Configuration invalid aggregate
    _bTimeout    : BOOL;                        // 建立超时保持量 / Held timeout value
    _bAging      : BOOL;                        // 老化预警保持量 / Held ageing warning
    _bInjectFault : BOOL;                       // 注入件故障 / Injected component fault
    _bVacReached : BOOL;                        // 真空已达目标 / Vacuum reached the target
    _bSampleNew  : BOOL;                        // 本次已入样本（单拍）/ A sample was buffered this scan
    _bBuildBrk   : BOOL := TRUE;                // 建立计时断输入一拍 / One-scan build break
    _bHeartBrk   : BOOL := TRUE;                // 心跳窗断输入一拍 / One-scan heartbeat break
    _nBaseUse    : INT;                         // 生效基线样本数，已钳制 [个] / Effective baseline sample count
    _nFill       : INT;                         // 已填样本数 [个] / Filled samples
    _nWriteIdx   : INT;                         // 环形写指针 [索引] / Ring write index
    _nWarnCnt    : INT;                         // 连续超门限计数 [次] / Consecutive exceed counter
    _nSortIdx    : INT;                         // 排序循环索引 [索引] / Sorting loop index
    _fSample     : ARRAY[0..15] OF REAL;        // 样本缓冲（建立时长）[ms] / Sample buffer [ms]
    _fMed        : REAL;                        // 中值 [ms] / Median [ms]
    _fBase       : REAL;                        // 基线保持量 [ms] / Held baseline [ms]
    _fDrift      : REAL;                        // 漂移保持量 [%] / Held drift [%]
    _fDevDen     : REAL;                        // 漂移分母（下限保护）[ms] / Drift denominator with a floor [ms]
    _fSortKey    : REAL;                        // 排序临时量（保留字，未参与秩计数法）[ms] / Sorting scratch reserved
    _nJ          : INT;                         // 内层循环索引 [索引] / Inner loop index
    _nRank       : INT;                         // 秩计数（严格小于本点的样本数）[个] / Rank counter
END_VAR
VAR CONSTANT
    DL_BASE_MAX   : INT := 16;          // 样本缓冲声明长度 [个] / Declared sample buffer length
    DL_MIN_SAMPLES : INT := 3;          // 出漂移结论的最少样本数 [个] / Minimum samples before a verdict
    DL_MS_FLOOR   : REAL := 1.0;        // 时长下限保护 [ms] / Duration floor to avoid division by zero
    DL_DRIFT_CLAMP_PCT : REAL := 500.0; // 漂移限幅 [%] / Drift clamp [%]
    DL_VAC_LIM_KPA : REAL := 200.0;     // 真空有限性上限 [kPa] / Vacuum magnitude ceiling [kPa]
    DL_HEART_WINDOW : TIME := T#2S;     // 心跳观察窗 [ms]，自复位节拍 / Heartbeat window, self-resetting
END_VAR

(* —— 段 0：定时器与边缘检测无条件周期刷新（R182：调用语句不得置于 IF / CASE 内） —— *)
rtReset(CLK := bReset);                                          // 复位上升沿，每拍必调
rtPick(CLK := bPickStart);                                       // 取料上升沿，每拍必调
tonHeart(IN := (NOT tonHeart.Q) AND (NOT _bHeartBrk), PT := DL_HEART_WINDOW);  // 心跳窗自复位
_bHeartBrk := FALSE;                                             // 断输入拍在调用后自清
tonBuild(IN := (_eState = E_DL_VacBuildState.eBuilding) AND (NOT _bBuildBrk), PT := tBuildMax);  // 建立计时
_bBuildBrk := FALSE;                                             // 断输入拍在调用后自清

(* —— 段 1：单拍量预清零（样本 / 基线 / 计数不入清单，R187①） —— *)
_uInfo      := 16#0000_0000;   // 信息码每拍重算
bError      := FALSE;          // 故障出口每拍重算，段 7 由锁存派生
bValid      := FALSE;          // 可用标志缺省 FALSE
_bCfgBad    := FALSE;          // 组态非法预清零
_bSampleNew := FALSE;          // 入样本单拍标志预清零
_bVacReached := FALSE;         // 真空达标判据预清零

(* —— 段 2：复位沿清锁存与保持量（R188 双路径） —— *)
IF rtReset.Q THEN
    _bFault   := FALSE;            // 复位沿清锁存位
    _uFault   := 16#0000_0000;     // 复位沿清锁存码
    _bTimeout := FALSE;            // 清建立超时保持量
    _bAging   := FALSE;            // 清老化预警保持量
    _nWarnCnt := 0;                // 清连续超门限计数
END_IF
IF (_uFault = 16#0003_0220) AND (NOT _bTimeout) THEN
    _uFault := 16#0000_0000;       // 按码专清：超时保持量已释放 → 对应码清除
    _bFault := FALSE;              // 锁存位同步清
END_IF

(* —— 段 3：组态域闸（覆盖全部参与换算的引脚，R151） —— *)
IF (fVacTargetKpa <> fVacTargetKpa) OR (fVacTargetKpa <= 0.0) OR (fVacTargetKpa > DL_VAC_LIM_KPA) THEN
    _bCfgBad := TRUE;              // 真空目标非法（建立判据门限）
END_IF
IF TIME_TO_DINT(tBuildMax) <= 0 THEN
    _bCfgBad := TRUE;              // 建立上限非法
END_IF
IF (fDriftWarnPct <> fDriftWarnPct) OR (fDriftWarnPct <= 0.0) THEN
    _bCfgBad := TRUE;              // 漂移门限非法
END_IF
IF nWarnCycles < 1 THEN
    _bCfgBad := TRUE;              // 连续次数门限非法
END_IF
_nBaseUse := nBaselineSamples;     // 生效样本数初值
IF _nBaseUse > DL_BASE_MAX THEN
    _nBaseUse := DL_BASE_MAX;      // 上限钳制（不静默截断，置信息码 0110）
    _uInfo := 16#0003_0110;        // 信息级：样本数超缓冲上限已钳制
END_IF
IF _nBaseUse < DL_MIN_SAMPLES THEN
    _nBaseUse := DL_MIN_SAMPLES;   // 下限钳制：低于 3 无中值意义
    _uInfo := 16#0003_0110;        // 信息级：样本数过小已抬升至最小可用值
END_IF
IF _bCfgBad THEN
    _uFault := 16#0003_0210;       // 故障级：组态非法
    _bFault := TRUE;               // 锁存位置位（复位沿可清）
    bError  := TRUE;               // 故障标志置位（R45 配对）
    _eState := E_DL_VacBuildState.eFault;  // 进故障相
END_IF

(* —— 段 4：真空反馈判据与注入件故障归因 —— *)
_bInjectFault := iVac.bFault;                                  // 注入件故障（不参与老化归因）
_bVacReached := ABS(iVac.fPressure) >= fVacTargetKpa;          // 真空达标（负压绝对值，分母无）
IF ABS(iVac.fPressure) > DL_VAC_LIM_KPA THEN
    _bCfgBad := TRUE;                                          // 真空反馈非有限/超上界：判据不可信
    _uFault := 16#0003_0210;                                   // 故障级：输入异常归入组态/输入异常码
    _bFault := TRUE;                                           // 锁存
    bError  := TRUE;                                           // 故障标志置位（R45 配对）
    _eState := E_DL_VacBuildState.eFault;                      // 进故障相
    _bVacReached := FALSE;                                     // 坏值不得当作达标
END_IF

(* —— 段 5：相位机（只做迁移与样本入缓冲；出口在段 8） —— *)
CASE _eState OF

E_DL_VacBuildState.eIdle:
    IF rtPick.Q AND bEnable AND (NOT _bFault) AND (NOT _bCfgBad) THEN
        _eState := E_DL_VacBuildState.eBuilding;          // 取料触发：进建立相
        _bBuildBrk := TRUE;                               // 建立计时从零
    END_IF

E_DL_VacBuildState.eBuilding:
    IF (NOT bEnable) THEN
        _eState := E_DL_VacBuildState.eIdle;              // 失能：放弃本次测量
    ELSIF _bVacReached THEN
        fBuildTimeMs := TIME_TO_REAL(tonBuild.ET);        // 本次建立时长 [ms]
        IF fBuildTimeMs < DL_MS_FLOOR THEN
            fBuildTimeMs := DL_MS_FLOOR;                  // 下限保护（同拍达成时不出现 0 时长）
        END_IF
        _fSample[_nWriteIdx] := fBuildTimeMs;             // 入环形样本缓冲
        _nWriteIdx := (_nWriteIdx + 1) MOD DL_BASE_MAX;   // 写指针推进（移位量已归一）
        IF _nFill < DL_BASE_MAX THEN
            _nFill := _nFill + 1;                         // 已填样本数饱和到缓冲长度
        END_IF
        _bSampleNew := TRUE;                              // 本拍已入样本（单拍）
        _bTimeout := FALSE;                               // 建立成功：超时保持量释放（按码专清的另一条边）
        _eState := E_DL_VacBuildState.eMeasured;          // 进已测量相
    ELSIF tonBuild.Q THEN
        _bTimeout := TRUE;                                // 建立超时保持量
        _uFault := 16#0003_0220;                          // 故障级：真空建立超时
        _bFault := TRUE;                                  // 锁存
        bError  := TRUE;                                  // 故障标志置位（R45 配对）
        _eState := E_DL_VacBuildState.eFault;             // 进故障相
    END_IF

E_DL_VacBuildState.eMeasured:
    IF (NOT bEnable) THEN
        _eState := E_DL_VacBuildState.eIdle;              // 失能：回空闲
    ELSIF rtPick.Q THEN
        _eState := E_DL_VacBuildState.eBuilding;          // 下一次取料：直接进建立相
        _bBuildBrk := TRUE;                               // 建立计时从零
    ELSE
        _eState := E_DL_VacBuildState.eIdle;              // 本次已完成：回空闲等待
    END_IF

E_DL_VacBuildState.eFault:
    IF (NOT _bFault) AND (NOT _bCfgBad) AND bEnable THEN
        _eState := E_DL_VacBuildState.eIdle;              // 锁存已清且组态合法：回空闲
    END_IF

ELSE
    _uFault := 16#0003_0230;                              // 故障级：相位 ID 越界（枚举兜底）
    _bFault := TRUE;                                      // 锁存
    bError  := TRUE;                                      // 故障标志置位（R45 配对）
    _eState := E_DL_VacBuildState.eFault;                 // 强制回故障相
END_CASE

(* —— 段 6：基线与漂移估计（中值抗野值；样本不足不出结论） —— *)
IF _bSampleNew AND (_nFill >= DL_MIN_SAMPLES) THEN
    (* 中值用秩计数法：对每点统计「严格小于它的样本数」，秩等于 nFill/2 者即中值。
       两层循环上界均由 _nFill 钳制（<= DL_BASE_MAX），无越界、无浮点相等比较 *)
    _fMed := _fSample[0];                                  // 中值初值（_nFill >= 3 已由外条件保证）
    FOR _nSortIdx := 0 TO (_nFill - 1) DO
        _nRank := 0;                                       // 本点秩计数清零
        FOR _nJ := 0 TO (_nFill - 1) DO
            IF _fSample[_nJ] < _fSample[_nSortIdx] THEN
                _nRank := _nRank + 1;                      // 严格小于本点的样本数
            END_IF
        END_FOR
        IF _nRank = (_nFill / 2) THEN
            _fMed := _fSample[_nSortIdx];                  // 秩等于半数的点即中值
        END_IF
    END_FOR
    _fBase := _fMed;                                       // 基线更新为中值 [ms]
    _fDevDen := MAX(_fBase, DL_MS_FLOOR);                  // 分母下限保护 [ms]
    _fDrift := (fBuildTimeMs - _fBase) / _fDevDen * 100.0; // 漂移 [%]（分母已证 >= 1 ms）
    IF _fDrift > DL_DRIFT_CLAMP_PCT THEN
        _fDrift := DL_DRIFT_CLAMP_PCT;                     // 上行限幅
    END_IF
    IF _fDrift < -DL_DRIFT_CLAMP_PCT THEN
        _fDrift := -DL_DRIFT_CLAMP_PCT;                    // 下行限幅
    END_IF
    IF _bInjectFault THEN
        _uInfo := 16#0003_0140;                            // 信息级：注入件故障，漂移结论抑制
        _nWarnCnt := 0;                                    // 抑制期不计连续次数
    ELSIF _fDrift > fDriftWarnPct THEN
        _nWarnCnt := _nWarnCnt + 1;                        // 连续超门限计数
        IF _nWarnCnt >= nWarnCycles THEN
            _bAging := TRUE;                               // 老化预警成立（维护级）
            _uInfo := 16#0003_0130;                        // 信息级：吸盘老化预警
        END_IF
    ELSE
        _nWarnCnt := 0;                                    // 未超门限：连续计数归零
        _bAging := FALSE;                                  // 漂移回落到门限内即自行释放（维护级可逆）
    END_IF
ELSIF _nFill < DL_MIN_SAMPLES THEN
    _uInfo := 16#0003_0120;                                // 信息级：样本不足，本拍不出漂移结论
    _fDrift := 0.0;                                        // 无基线：漂移置 0（不产生 inf/NaN）
    _bAging := FALSE;                                      // 无结论：不置老化预警
END_IF

(* —— 段 7：故障码优先级链（每个 bError 置位源在此均有码，R45 配对） —— *)
IF _bCfgBad THEN
    _uFault := 16#0003_0210;                               // 组态非法优先上报
    _bFault := TRUE;
    bError  := TRUE;
END_IF

(* —— 段 8：出口单点映射（名实同源；锁存码回放，禁同拍抹除） —— *)
fBaselineMs   := _fBase;                                   // 基线出口 [ms]
fDriftPct     := _fDrift;                                  // 漂移出口 [%]
bAgingWarn    := _bAging AND (NOT _bInjectFault);          // 老化预警出口（注入件故障期抑制）
bBuildTimeout := _bTimeout;                                // 建立超时出口（保持型）
nSampleCount  := _nFill;                                   // 有效样本数出口
eStateOut     := _eState;                                  // 状态出口
IF _bFault THEN
    nErrId := _uFault;                                     // 故障锁存码回放（不在故障相按当下输入重推）
    bError := TRUE;                                        // 故障出口派生自锁存
ELSE
    nErrId := _uInfo;                                      // 信息码
END_IF
bValid := bEnable AND (NOT _bFault) AND (NOT _bCfgBad);    // 判据可用

END_FUNCTION_BLOCK
